(* IEC 61131-3 sources: daoli-st-library/DL_Process (part 57) *)

(* ---- FB_DL_TrapSealTrend.st ---- *)
(*
  FB_DL_TrapSealTrend  —  枕式包装封口温度随线速前馈重置 / Pillow-pack seal temperature feedforward with line-speed reset
  分类 Category : DL_Process
  码位 Code     : 16#06_0_86
  版本 Version  : 1.0.1
  溯源 Source   : Modular PID 语义借鉴 · clean-room 实现，仅借分类/参数域/命名，未复制源码
  修订 Revision : v1.0.1 (R34 终审抽检) — ① 判停改按原始线速 bSpeedStop，修正「零速保持相在曾运行后不可达」
                  （原以 fSpeedUse 判停，而 fSpeedUse 是末次有效线速替代值，恒 > 0 致 bHold 永假）；
                  ② 输入引脚 fSpeedValid 更名 bSpeedValid（BOOL 前缀红线 1，v1.0.0 无下游调用方，不构成破坏性变更）；
                  ③ 删段 7 自赋值空语句 uInfo := uInfo。接口语义与码表不变。
  功能 Function : 1) 线速前馈：封温设定 = 基准设定 + 线速偏差 × 前馈增益，线速经斜坡限速后进 PID 设定；
                  2) 线速为 0 时不得外推封温设定，改用末次有效线速并置 bHold（禁按零速反推冷设定）；
                  3) 封温设定钳到工艺窗口上下限，越限只钳位 + 报码不拒算；重置斜率须与 PID 采样周期配比，超调即判组态非法。
  边界 Boundary : ① 线速为 0 不得外推封温设定（末次有效线速 + bHold）；
                  ② 重置限速斜率与 PID 采样周期配比（每采样步进 <= fSpStepMaxC），非法即组态报码；
                  ③ 封温设定钳到工艺窗口上下限，越限只钳位 + 报码不拒算；
                  ④ 安全侧三行同向：PID 输出限 0 → 设定保持末值 → bHold 置位。
  依赖 Depends  : FB_DL_PidController（封温闭环）、FB_DL_RateLimiter（设定斜坡），均每拍无条件调用

  码表 Error codes（本件子码步进 16#10，避让邻件码位）:
    16#0002_0686 故障级：组态非法（工艺窗口上/下限倒置、增益或斜率 <= 0、采样周期 <= 0）
    16#0002_0696 故障级：前馈斜率与采样周期配比超调（单步进料过大）
    16#0002_06A6 信息级：封温设定已钳位（不置 bError，照算）
*)

TYPE E_DL_TstPhase :
(
    eIdle   := 0,   // 空闲 / Idle
    eTrack  := 10,  // 线速跟踪 / Line-speed tracking
    eHold   := 20,  // 零速保持 / Zero-speed hold
    eRun    := 30,  // 闭环调节 / Closed-loop control
    eFault  := 90   // 故障锁定 / Fault locked
);
END_TYPE

FUNCTION_BLOCK FB_DL_TrapSealTrend
VAR_INPUT
    bEnable      : BOOL;                          // 总使能，FALSE 回空闲 / Master enable
    bReset       : BOOL;                          // 复位，上升沿清故障 / Reset, clears fault
    fLineSpeedMpm: REAL;                          // 包装线速 [m/min]，域 >= 0 / Packaging line speed [m/min]
    bSpeedValid  : BOOL := TRUE;                  // 线速信号有效标志 / Line speed signal valid
    fSealTempC   : REAL;                          // 封口实测温度 [degC]，域 0~300 / Measured seal temperature [degC]
    fSealBaseC   : REAL := 150.0;                 // 基准封温设定 [degC] / Base seal temperature setpoint [degC]
    fFfGainCpm   : REAL := 0.8;                   // 线速前馈增益 [degC per m/min]，域 > 0 / Feedforward gain
    fSealWinLoC  : REAL := 120.0;                 // 工艺窗口下限 [degC] / Process window low [degC]
    fSealWinHiC  : REAL := 200.0;                 // 工艺窗口上限 [degC] / Process window high [degC]
    fSpRiseRate  : REAL := 20.0;                  // 设定上升限速 [degC/s]，域 > 0 / Setpoint rise rate [degC/s]
    fSpFallRate  : REAL := 20.0;                  // 设定下降限速 [degC/s]，域 > 0 / Setpoint fall rate [degC/s]
    fSpStepMaxC  : REAL := 5.0;                   // 单采样步进上限 [degC]，域 > 0 / Step limit per sample [degC]
    tPidSample   : TIME := T#100MS;               // PID 采样周期 [ms]，域 > 0 / PID sample period [ms]
    fKp          : REAL := 2.0;                   // 比例增益 [1] / Proportional gain
    tTi          : TIME := T#30S;                 // 积分时间 [ms] / Integral time [ms]
    tTd          : TIME := T#5S;                  // 微分时间 [ms] / Derivative time [ms]
    fEps         : REAL := 1.0E-6;                // 浮点判零容差 [1] / Floating zero tolerance
END_VAR
VAR_OUTPUT
    fSealSpC     : REAL;                          // 封温设定 [degC]，经前馈 + 限速 + 钳位 / Seal setpoint [degC]
    fPidOutPct   : REAL;                          // 加热输出 [%] / Heater output [%]
    fSpeedHold   : REAL;                          // 生效线速 [m/min]，零速时保持末次有效 / Effective line speed
    bHold        : BOOL;                          // 零速保持标志 / Zero-speed hold flag
    bClamped     : BOOL;                          // 设定钳位标志 / Setpoint clamped flag
    bError       : BOOL;                          // 故障标志，与故障级码配对 / Fault flag paired with fault codes
    uErrorId     : UDINT;                         // 事件码，0 = 无事件 / Event code, 0 = none
    eStateOut    : E_DL_TstPhase;                 // 状态机当前态，段尾单点映射 / Phase mapped at tail
END_VAR
VAR
    _eState      : E_DL_TstPhase := E_DL_TstPhase.eIdle;  // 内部状态 / Internal state
    rtrReset     : R_TRIG;                        // 复位沿 / Reset edge
    fbPid        : FB_DL_PidController;           // 封温闭环实例（无条件调用）/ Seal loop PID
    fbSpRamp     : FB_DL_RateLimiter;             // 设定斜坡实例（无条件调用）/ Setpoint ramp limiter
    bCfgOk       : BOOL;                          // 组态合法标志 / Configuration valid
    bRatioOk     : BOOL;                          // 斜率/周期配比合法 / Slope-period ratio valid
    fSpeedUse    : REAL;                          // 前馈用线速 [m/min] / Speed used for feedforward
    bSpeedStop   : BOOL;                          // 线速判停标志（按原始线速判，非替代值）/ Line stopped per raw speed
    fSpRawC      : REAL;                          // 前馈原始设定 [degC] / Raw feedforward setpoint [degC]
    fSampleS     : REAL;                          // 采样周期折算秒 [s] / Sample period in seconds
    fStepC       : REAL;                          // 单采样最大步进 [degC] / Max step per sample [degC]
    uFault       : UDINT;                         // 锁存故障码 / Latched fault code
    uInfo        : UDINT;                         // 信息级码 / Information code
END_VAR
VAR CONSTANT
    DL_TST_MSPS    : REAL := 1000.0;              // 毫秒折算秒系数 [ms/s] / Milliseconds per second
    DL_TST_TMAXC   : REAL := 300.0;               // 封温物理域上限 [degC] / Temperature domain high
END_VAR

(* === 段 0 · 实例刷新（无条件周期调用，禁入 CASE 分支）=== *)
rtrReset(CLK := bReset);                          // 每拍刷新复位沿

(* === 段 1 · 组态闸：窗口配比 / 增益正域 / 斜率-周期配比 === *)
fSampleS := TIME_TO_LREAL(tPidSample) / DL_TST_MSPS;   // 采样周期折算秒，标准转换函数
bCfgOk := (fSealWinHiC > fSealWinLoC) AND (fFfGainCpm > fEps) AND (fSpRiseRate > fEps)
          AND (fSpFallRate > fEps) AND (fSpStepMaxC > fEps) AND (fSampleS > fEps)
          AND (fSealBaseC > 0.0) AND (fSealBaseC < DL_TST_TMAXC)
          AND (fSealWinHiC = fSealWinHiC) AND (fSealWinLoC = fSealWinLoC);   // NaN 自反判据
fStepC := fSpRiseRate * fSampleS;                 // 单采样步进 = 斜率 × 周期
bRatioOk := (fStepC <= fSpStepMaxC + fEps);       // 配比闸：单步进不得超过工艺允许步进（超调即非法）
IF NOT bCfgOk THEN
    uFault := 16#0002_0686;                       // 故障级：组态非法
END_IF
IF NOT bRatioOk THEN
    uFault := 16#0002_0696;                       // 故障级：斜率与采样周期配比超调
END_IF
IF rtrReset.Q AND bCfgOk AND bRatioOk THEN
    uFault := 16#0000;                            // 复位沿清锁存（故障复位路径可达）
END_IF
uInfo := 16#0000;                                 // 信息码每拍清零

(* === 段 2 · 线速域闸：零速/无效速保持末次有效，不外推 === *)
bSpeedStop := (NOT bSpeedValid) OR (fLineSpeedMpm <> fLineSpeedMpm) OR (fLineSpeedMpm <= fEps);  // 判停只看原始线速（NaN 自反捕获）
IF NOT bSpeedStop
   AND (ABS(fLineSpeedMpm) < 1.0E6) THEN
    fSpeedUse := fLineSpeedMpm;                   // 有效线速直接采用
    fSpeedHold := fLineSpeedMpm;                  // 记入末次有效线速
ELSE
    fSpeedUse := fSpeedHold;                      // 零速/无效：用末次有效线速，禁按 0 反推
END_IF
fSpRawC := fSealBaseC + fSpeedUse * fFfGainCpm;   // 前馈原始设定 [degC]

(* === 段 3 · 设定斜坡实例（每拍无条件调用，限斜率）=== *)
fbSpRamp(bEnable := TRUE,                         // 斜坡常开
         fIn := fSpRawC,                          // 前馈原始设定
         fRateUp := fSpRiseRate,                  // 上升限速 [degC/s]
         fRateDown := fSpFallRate,                // 下降限速 [degC/s]
         bTrack := (NOT bEnable) OR (uFault <> 16#0000),   // 失能/故障：跟踪到基准设定
         fTrackValue := fSealBaseC,               // 跟踪目标 = 基准设定
         tSampleTime := tPidSample);              // 采样周期
fSealSpC := fbSpRamp.fOut;                        // 斜坡后设定

(* === 段 4 · 封温窗口钳位（越限只钳位 + 报码，不拒算）=== *)
bClamped := FALSE;                                // 钳位标志每拍重算
IF fSealSpC > fSealWinHiC THEN
    fSealSpC := fSealWinHiC;                      // 钳到上限
    bClamped := TRUE;                             // 钳位置位
    uInfo := 16#0002_06A6;                        // 信息级：设定已钳位
ELSIF fSealSpC < fSealWinLoC THEN
    fSealSpC := fSealWinLoC;                      // 钳到下限
    bClamped := TRUE;                             // 钳位置位
    uInfo := 16#0002_06A6;                        // 信息级：设定已钳位
END_IF

(* === 段 5 · 主状态机（ENUM + CASE，含 ELSE 兜底）=== *)
CASE _eState OF
E_DL_TstPhase.eIdle :
    bHold := FALSE;                               // 空闲不保持
    IF uFault <> 16#0000 THEN
        _eState := E_DL_TstPhase.eFault;          // 故障优先
    ELSIF bEnable THEN
        _eState := E_DL_TstPhase.eTrack;          // 进入跟踪相
    END_IF

E_DL_TstPhase.eTrack :
    IF bSpeedStop THEN                            // 判停按原始线速（不按前馈替代值）
        bHold := TRUE;                            // 零速：置保持，禁止外推冷设定
        _eState := E_DL_TstPhase.eHold;
    ELSE
        bHold := FALSE;                           // 有速：正常调节
        _eState := E_DL_TstPhase.eRun;
    END_IF

E_DL_TstPhase.eHold :
    bHold := TRUE;                              // 保持标志维持
    IF NOT bSpeedStop THEN
        bHold := FALSE;                          // 线速恢复即解除保持（可到达的解除路径）
        _eState := E_DL_TstPhase.eRun;
    END_IF

E_DL_TstPhase.eRun :
    IF bSpeedStop THEN                           // 判停按原始线速，与 eTrack 同源
        bHold := TRUE;                            // 线速降到 0：回保持
        _eState := E_DL_TstPhase.eHold;
    ELSIF NOT bEnable THEN
        _eState := E_DL_TstPhase.eIdle;           // 失能回空闲
    ELSIF uFault <> 16#0000 THEN
        _eState := E_DL_TstPhase.eFault;          // 故障拦截
    END_IF

E_DL_TstPhase.eFault :
    bHold := TRUE;                                // 故障态保持（安全侧）
    IF uFault = 16#0000 THEN
        _eState := E_DL_TstPhase.eIdle;           // 解锁回空闲
    END_IF

ELSE
    _eState := E_DL_TstPhase.eFault;              // 非法状态拦截
    uFault := 16#0002_0686;                       // 故障级：相 ID 越界（枚举兜底路径）
END_CASE

(* === 段 6 · 封温闭环实例（每拍无条件调用）=== *)
fbPid(bEnable := bEnable AND (NOT bHold) AND (uFault = 16#0000),   // 保持/故障时禁调节
      bManual := FALSE,                           // 自动模式
      fManualValue := 0.0,                        // 手动值未用
      fSetpoint := fSealSpC,                      // 设定 = 钳位后封温
      fActual := fSealTempC,                      // 实测封温
      fKp := fKp,                                 // 比例增益
      tTi := tTi,                                 // 积分时间
      tTd := tTd,                                 // 微分时间
      fDeadband := 0.5,                           // 控制死区 [degC]，防抖
      bIncremental := FALSE,                      // 位置式
      rOutMin := 0.0,                             // 输出下限 0%（安全侧）
      rOutMax := 100.0,                           // 输出上限 100%
      tSampleTime := tPidSample,                  // 采样周期
      bTrack := bHold OR (uFault <> 16#0000),     // 保持/故障：跟踪 0 输出
      fTrackValue := 0.0,                         // 跟踪值 0（断加热）
      bReset := rtrReset.Q);                      // 复位沿清积分

(* === 段 7 · 输出映射（安全三行同向）=== *)
IF bHold OR (uFault <> 16#0000) THEN
    fPidOutPct := 0.0;                            // 保持/故障：加热输出 0（驱动方向安全）
    bHold := TRUE;                                // 保持判据与输出同向（设定同步冻结在段 3/4 末值）
ELSE
    fPidOutPct := fbPid.fOut;                     // 正常：取 PID 输出
END_IF
IF NOT bEnable THEN
    fPidOutPct := 0.0;                            // 失能输出 0
END_IF
bError := (uFault <> 16#0000);                    // 故障标志仅由故障级码置位（R45 配对）
IF bError THEN
    uErrorId := uFault;                           // 故障级优先上报
ELSE
    uErrorId := uInfo;                            // 否则上报信息级码
END_IF
eStateOut := _eState;                             // 输出枚举段尾单点映射（N2 规则）
END_FUNCTION_BLOCK

(* ---- FB_DL_TrayerNestingCtrl.st ---- *)
(*==============================================================================
 * 组件名称 (Component)  : FB_DL_TrayerNestingCtrl
 * 所属子库 (Sublibrary) : DL_Process
 * 当前版本 (Version)    : 1.0.0
 * 兼容性   (Platform)   : CODESYS 3.5+ / TwinCAT 3 / 汇川 InoProShop / 施耐德 Machine Expert
 *                         仅依赖 Standard.library（R_TRIG），零厂商私有库
 * 功能描述 (Function)   : 电芯托盘堆叠嵌套调度（层 × 列网格占位）。
 *                         按"层从下往上、列从左往右"的蛇形无关直线序逐格占位；每来一颗电芯占一格，
 *                         列到边界回卷到下一层首列；**NG 通道避让**：某一列指定为 NG 列时，
 *                         该列在每一层都被整体跳过（整列不占位、不计入容量）；
 *                         合法格占满即判"栈满"并锁存 bTrayFull，等待取盘沿（bTrayTaken）或复位沿解除。
 *                         **语义复用（非实例复用）**：本件按 R47 批次"批内零 .st 文件级依赖"纪律，
 *                         不实例化 FB_DL_LifoStack，而是复用其三条已固化语义——
 *                         ① 入栈前判满、满则拒入并锁存；② 出栈仅由显式"取走"沿触发；
 *                         ③ 满/空判定以计数与容量比较为准，不以指针相等为准。
 *                         验收向量：
 *                           ① 3 层 × 4 列、NG 列 = 2 → 容量 = 3×(4−1) = 9 格
 *                           ② 2 层 × 2 列、NG 列 = 1 → 容量 = 2×(2−1) = 2 格
 *                           ③ 2 层 × 2 列、NG 列 = 0 → 容量 = 4 格
 *                           ④ 任一层列数 = 0 → 组态非法锁存，不进入占位
 * 接口     (Interface)  : 入 bStart 启动沿、bTrayTaken 取盘沿（解除栈满）、iLayerCnt 层数、iColCnt 列数、
 *                         iNgCol 避让列号（1 基，0 = 无）、bCellPresent 电芯到位沿、bPlaceAllowed 上料允许
 *                         （外部互锁）、bReset 故障复位沿；
 *                         出 iLayerOut / iColOut 当前待占格坐标（1 基）、bPlaceCmd 占位脉冲（单拍）、
 *                         bLayerDone 换层脉冲（单拍）、bTrayFull 栈满锁存、iPlacedCnt 已占格数、
 *                         bNgSkipped 当拍发生 NG 列跳过、eState 相、eCause 成因、bError 故障标志。
 * 边界     (Boundary)   : ① **属主边界（写死）：本件只算"下一颗电芯放哪一格"，不驱动吸盘/夹具/
 *                         升降台伺服**；取放动作由执行件（I_DL_Cylinder 族 / 运动件）承担；
 *                         ② **网格组态闸**：层数或列数 ≤ 0 或超上限（100×100）→ 锁存 eCfgIllegal，
 *                         不进入占位（零容量网格会让"栈满"永假，属静默失效 R179）；
 *                         ③ **NG 列域闸**：iNgCol 越界（<0 或 > 列数）→ 锁存 eCfgIllegal；
 *                         ④ **索引越界钳位**：前进循环带 _uGuard 计数器（上界 = 总格数 + 列数 + 2），
 *                         循环必然收敛，绝不靠"数据一定合法"保证终止；
 *                         ⑤ eFault 可迁出：bReset 上升沿 → eIdle（解除式自证：bReset 为外部引脚，
 *                         不受任何锁存量门控，恒可达）；
 *                         ⑥ 零全局耦合、零物理地址。
 * 分工声明 (Scope)      : 本件只管"托盘格位调度与栈满判定"。不接管：电芯取放动作时序（顺控件）、
 *                         NG 电芯的下游分选（分选件）、托盘身份绑定（RFID 件）。
 * 来源标签 (Source Tag) : ROADMAP 空勾真缺口 P2（托盘嵌套调度，自研 clean-room）
 * 码表     (Codes)      : 本件不占用任何全局数字码位（零码位范式 R297）；诊断由 BOOL + ENUM 出口承担。
 * 红线自检 (Redline)    : R1 ✓ 零 GVL/VAR_EXTERNAL ｜ R2 ✓ 零 %I/%Q/%M ｜ R3 ✓ 纯 IEC 61131-3
 *                         R4 ✓ 组态双闸 + 循环计数器 + 索引钳位 ｜ R5 ✓ 声明逐行同行双语注释
 *                         R6 ✓ ENUM+CASE 含 ELSE 兜底 ｜ R7 ✓ R_TRIG 段 0 无条件刷新（本件无 TON）
 * 修订历史 (Revision)   : 2026-11-19  v1.0.0  R47 首版（批次 1 · 序号 4）
 *==============================================================================*)

TYPE E_DL_TncState :
(
    eIdle  := 0,    // 待机相（等启动或等取盘） / Idle, awaiting start or tray removal
    eNest  := 10,   // 占位相（逐颗占格） / Nesting, one cell per cell-in
    eFull  := 20,   // 栈满相（锁存等取盘） / Full, latched awaiting tray removal
    eFault := 90    // 故障相（等复位） / Fault, awaiting reset
);
END_TYPE

TYPE E_DL_TncCause :
(
    eNone      := 0,   // 无异常 / No anomaly
    eCfgIllegal:= 1,   // 组态非法（层数/列数/NG 列越域） / Illegal grid configuration
    eFullNoCell    := 2,   // 栈满后仍有电芯到位（拒入） / Cell arrived while full, rejected
    eRejectNoPermit:= 3,   // 上料允许缺失致电芯被拒 / Cell rejected, place permit absent
    ePhaseBad      := 4    // 非法相位兜底 / Illegal phase fallback
);
END_TYPE

FUNCTION_BLOCK FB_DL_TrayerNestingCtrl
VAR_INPUT
    bStart       : BOOL := FALSE;   // 启动沿，进入占位相 [-] / Start edge, enters nesting
    bTrayTaken   : BOOL := FALSE;   // 取盘沿，解除栈满并清零计数 [-] / Tray-removed edge, clears the full latch
    iLayerCnt    : INT := 1;        // 层数，域 1..100 [层] / Layer count, domain 1..100
    iColCnt      : INT := 1;        // 每层列数，域 1..100 [列] / Columns per layer, domain 1..100
    iNgCol       : INT := 0;        // NG 避让列号（1 基；0 = 不避让） [列] / NG column index, 1-based, 0 = none
    bCellPresent : BOOL := FALSE;   // 电芯到位信号（上升沿占一格） [-] / Cell-present signal, rising edge takes one cell
    bPlaceAllowed: BOOL := FALSE;   // 上料允许（外部互锁，FALSE 时拒占位） [-] / Place permit from the external interlock
    bReset       : BOOL := FALSE;   // 故障复位沿 [-] / Fault reset edge
END_VAR
VAR_OUTPUT
    iLayerOut  : INT := 0;                  // 当前待占格所在层（1 基） [层] / Current target layer, 1-based
    iColOut    : INT := 0;                  // 当前待占格所在列（1 基） [列] / Current target column, 1-based
    bPlaceCmd  : BOOL := FALSE;             // 占位脉冲，单拍 [-] / Place command, single-scan pulse
    bLayerDone : BOOL := FALSE;             // 换层脉冲，单拍 [-] / Layer-change pulse, single-scan
    bTrayFull  : BOOL := FALSE;             // 栈满锁存（等取盘或复位） [-] / Tray full, latched
    iPlacedCnt : INT := 0;                  // 已占格数 [格] / Occupied cell count
    bNgSkipped : BOOL := FALSE;             // 当拍发生过 NG 列跳过 [-] / An NG column was skipped this scan
    eState     : E_DL_TncState := E_DL_TncState.eIdle;   // 相出口 [-] / Phase outlet
    eCause     : E_DL_TncCause := E_DL_TncCause.eNone;   // 成因出口（R190 归因唯一） [-] / Cause outlet
    bError     : BOOL := FALSE;             // 故障标志 [-] / Error flag
END_VAR
VAR
    _eState    : E_DL_TncState := E_DL_TncState.eIdle;   // 内部相（CASE 唯一写入目标） / Internal phase
    _eCause    : E_DL_TncCause := E_DL_TncCause.eNone;   // 成因锁存量 / Latched cause
    _bFault    : BOOL := FALSE;             // 故障锁存位 / Latched fault bit
    _bFull     : BOOL := FALSE;             // 栈满锁存位（与 bTrayFull 同源） / Latched full bit
    _iLayer    : INT := 1;                  // 内部层指针（1 基） / Internal layer cursor
    _iCol      : INT := 1;                  // 内部列指针（1 基） / Internal column cursor
    _iPlaced   : INT := 0;                  // 内部已占格计数 / Internal occupied counter
    _iCap      : INT := 0;                  // 本盘合法格容量（不含 NG 列） / Legal capacity excluding the NG column
    _bPlaceCmd : BOOL := FALSE;             // 占位脉冲内部位（单拍） / Internal place pulse
    _bLayerDone: BOOL := FALSE;             // 换层脉冲内部位（单拍） / Internal layer-change pulse
    _bNgSkipped: BOOL := FALSE;             // NG 跳过内部位（单拍） / Internal NG-skip flag
    _bCfgBad   : BOOL := FALSE;             // 组态非法当拍量 / Illegal configuration this scan
    _bAdvDone  : BOOL := FALSE;             // 前进循环收敛标志 / Advance-loop convergence flag
    _uGuard    : UINT := 0;                 // 前进循环计数器（防死循环） / Advance-loop guard counter
    rtStart    : R_TRIG;                    // 启动沿实例，段 0 无条件调用 / Start edge instance
    rtReset    : R_TRIG;                    // 复位沿实例，段 0 无条件调用 / Reset edge instance
    rtTaken    : R_TRIG;                    // 取盘沿实例，段 0 无条件调用 / Tray-removed edge instance
    rtCell     : R_TRIG;                    // 电芯到位沿实例，段 0 无条件调用 / Cell-present edge instance
END_VAR
VAR CONSTANT
    DL_TNC_MAX_LAYER : INT := 100;          // 层数上限（超限判组态非法） [层] / Layer upper bound
    DL_TNC_MAX_COL   : INT := 100;          // 列数上限（超限判组态非法） [列] / Column upper bound
    DL_TNC_GUARD_MAX : UINT := 20002;       // 前进循环守护上限（100×100 + 100 + 2） [次] / Advance guard limit
END_VAR

(* —— 段 0：组态闸 + 四枚沿实例无条件周期刷新（R228A） —— *)
_bCfgBad := (iLayerCnt <= 0) OR (iLayerCnt > DL_TNC_MAX_LAYER)          // 层数须在 1..100 / Layer count within 1..100
         OR (iColCnt <= 0) OR (iColCnt > DL_TNC_MAX_COL)                // 列数须在 1..100 / Column count within 1..100
         OR (iNgCol < 0) OR (iNgCol > iColCnt);                          // NG 列号须为 0 或落在列域内 / NG index within the column domain
rtStart(CLK := bStart);                                                  // 启动沿 / Start edge
rtReset(CLK := bReset);                                                  // 复位沿 / Reset edge
rtTaken(CLK := bTrayTaken);                                              // 取盘沿 / Tray-removed edge
rtCell(CLK := bCellPresent);                                             // 电芯到位沿 / Cell-present edge

(* —— 段 1：单拍量预清零（锁存量 _eCause/_bFault/_iPlaced 不入清单，R107） —— *)
_bPlaceCmd  := FALSE;                                                    // 占位脉冲预清 / Place pulse preset
_bLayerDone := FALSE;                                                    // 换层脉冲预清 / Layer pulse preset
_bNgSkipped := FALSE;                                                    // NG 跳过标志预清 / NG-skip preset
bError      := FALSE;                                                    // 故障标志预清（R45 配对） / Error preset

(* —— 段 2：组态闸（非法即锁存，不进入占位） —— *)
IF _bCfgBad THEN
    _bFault := TRUE;                                                     // 锁存 / Latch
    _eCause := E_DL_TncCause.eCfgIllegal;                                // 归因：组态非法 / Cause: illegal configuration
    _eState := E_DL_TncState.eFault;                                     // 入故障相 / Enter fault phase
END_IF

(* —— 段 3：迁出链与取盘链（两条出口显式写出，R228B） —— *)
IF rtReset.Q THEN
    _bFault  := FALSE;                                                   // 清故障锁存 / Clear fault latch
    _bFull   := FALSE;                                                   // 清栈满锁存 / Clear full latch
    _eCause  := E_DL_TncCause.eNone;                                     // 清成因 / Clear cause
    _iPlaced := 0;                                                       // 计数清零 / Clear the counter
    _iLayer  := 1;                                                       // 层指针回 1 / Layer cursor back to 1
    _iCol    := 1;                                                       // 列指针回 1 / Column cursor back to 1
    _eState  := E_DL_TncState.eIdle;                                     // 回待机相 / Back to idle
END_IF
IF rtTaken.Q AND (_eState <> E_DL_TncState.eFault) THEN
    _bFull   := FALSE;                                                   // 取盘解除栈满 / Tray removal clears the full latch
    _iPlaced := 0;                                                       // 计数清零 / Clear the counter
    _iLayer  := 1;                                                       // 层指针回 1 / Layer cursor back to 1
    _iCol    := 1;                                                       // 列指针回 1 / Column cursor back to 1
    _eState  := E_DL_TncState.eIdle;                                     // 回待机相 / Back to idle
END_IF

(* —— 段 4：容量计算（总格数 − NG 列整列格数；组态合法时恒 ≥ 0） —— *)
IF NOT _bCfgBad THEN
    _iCap := iLayerCnt * iColCnt;                                        // 总格数 / Total cells
    IF iNgCol > 0 THEN
        _iCap := _iCap - iLayerCnt;                                      // 扣除 NG 列整列 / Deduct the whole NG column
    END_IF
END_IF

(* —— 段 5：相迁移（只在无故障时推进；每相出口条件显式成对） —— *)
IF (NOT _bFault) AND (NOT _bCfgBad) THEN
    CASE _eState OF

    E_DL_TncState.eIdle:
        IF rtStart.Q THEN
            _iLayer := 1;                                                // 层指针首层 / First layer
            IF (iNgCol = 1) AND (iColCnt >= 2) THEN
                _iCol := 2;                                              // 首列即 NG：起始列右移一格 / First column is NG, start at column 2
            ELSE
                _iCol := 1;                                              // 否则首列起步 / Otherwise start at column 1
            END_IF
            _iPlaced := 0;                                               // 计数清零 / Counter cleared
            _eState := E_DL_TncState.eNest;                              // 进占位相 / Enter nesting
        END_IF

    E_DL_TncState.eNest:
        IF rtCell.Q AND bPlaceAllowed THEN
            _bPlaceCmd := TRUE;                                          // 占位脉冲（内部位，段 7 单点映射） / Internal place pulse
            _iPlaced := _iPlaced + 1;                                    // 占位计数 +1 / Increment the counter

            (* 前进到下一合法格：列 +1，越界回卷到下一层首列，NG 列整体跳过 *)
            _uGuard  := 0;                                               // 守护计数器归零 / Guard reset
            _bAdvDone:= FALSE;                                           // 收敛标志复位 / Convergence flag reset
            WHILE (NOT _bAdvDone) AND (_uGuard < DL_TNC_GUARD_MAX) DO
                _uGuard := _uGuard + 1;                                  // 计数器推进 / Guard advance
                _iCol := _iCol + 1;                                      // 列前进一格 / Column step
                IF _iCol > iColCnt THEN
                    _iCol := 1;                                          // 列回卷 / Column wrap
                    _iLayer := _iLayer + 1;                              // 换层 / Next layer
                    _bLayerDone := TRUE;                                 // 换层脉冲（内部位） / Internal layer pulse
                END_IF
                IF _iLayer > iLayerCnt THEN
                    _bAdvDone := TRUE;                                   // 层耗尽：指针停（不再寻格） / Layers exhausted
                ELSIF (iNgCol > 0) AND (_iCol = iNgCol) THEN
                    _bNgSkipped := TRUE;                                 // NG 列：跳过并继续寻格 / NG column skipped, keep seeking
                ELSE
                    _bAdvDone := TRUE;                                   // 找到合法格 / Legal cell found
                END_IF
            END_WHILE

            IF _iPlaced >= _iCap THEN
                _bFull   := TRUE;                                        // 栈满锁存（入栈前判满语义） / Full latch, pre-push check
                _eState  := E_DL_TncState.eFull;                         // 进栈满相 / Enter full phase
            END_IF
        ELSIF rtCell.Q AND (NOT bPlaceAllowed) THEN
            _eCause := E_DL_TncCause.eRejectNoPermit;                    // 归因：互锁未放开致电芯被拒 / Cause: cell rejected, permit absent
        END_IF

    E_DL_TncState.eFull:
        IF rtCell.Q THEN
            _eCause := E_DL_TncCause.eFullNoCell;                        // 满盘期电芯到位：拒入并留痕 / Cell during full: rejected and recorded
        END_IF

    E_DL_TncState.eFault:
        ;                                                                // 故障相：由段 3 复位沿迁出 / Exit handled by the reset edge in stage 3

    ELSE
        _eCause := E_DL_TncCause.ePhaseBad;                              // 归因：非法相位 / Cause: illegal phase
        _bFault := TRUE;                                                 // 锁存 / Latch
        _eState := E_DL_TncState.eFault;                                 // 强拉故障相 / Force fault phase

    END_CASE
END_IF

(* —— 段 6：栈满与故障的交汇（满盘后故障优先展示，满锁存保持） —— *)
IF _bFull AND (_eState = E_DL_TncState.eNest) THEN
    _eState := E_DL_TncState.eFull;                                      // 满锁存与相对齐 / Align the phase with the full latch
END_IF

(* —— 段 7：出口单点映射（名实双出口，R191） —— *)
iLayerOut  := _iLayer;                                                   // 待占层层号 / Target layer
iColOut    := _iCol;                                                     // 待占格列号 / Target column
bPlaceCmd  := _bPlaceCmd;                                                // 占位脉冲单拍出口 / Place pulse outlet
bLayerDone := _bLayerDone;                                               // 换层脉冲单拍出口 / Layer pulse outlet
bNgSkipped := _bNgSkipped;                                               // NG 跳过标志出口 / NG-skip outlet
bTrayFull  := _bFull;                                                    // 栈满出口 / Full outlet
iPlacedCnt := _iPlaced;                                                  // 已占格数出口 / Occupied count outlet
eState     := _eState;                                                   // 相出口 / Phase outlet
eCause     := _eCause;                                                   // 成因出口 / Cause outlet
bError     := _bFault OR _bCfgBad;                                       // 故障标志 = 锁存或组态非法 / Error = latch or illegal config

END_FUNCTION_BLOCK

(* ---- FB_DL_TrayLoadVacuum.st ---- *)
(*==============================================================================
 * 组件名称 (Component)  : FB_DL_TrayLoadVacuum
 * 所属子库 (Sublibrary) : DL_Process
 * 当前版本 (Version)    : 1.0.0
 * 兼容性 (Platform)     : CODESYS 3.5+ / TwinCAT 3 / 汇川 InoProShop / 施耐德 Machine Expert
 *                         仅依赖 Standard.library（TON / TOF / R_TRIG / F_TRIG），零厂商私有库
 * 功能描述 (Function)   : 电池片花篮真空取放顺控。吸取相开真空阀，真空反馈
 *                         在 tVacOnDelay 内不到达即吸取超时故障（独立成因）；
 *                         放片相关真空并以 TOF 定宽输出破真空吹气脉冲
 *                         （宽度 tBlowWidth + 1 扫描拍，头注释明示），吹气
 *                         结束沿收口 bPlaceDone。与 VacuumEjector（真空发生
 *                         设备件）分工：本件是取放顺控中破真空定宽脉冲的
 *                         时序件。
 * 来源标签 (Origin)     : ROADMAP §9.3 P2（L418），自研 clean-room
 * 边界语义 (Boundary)   : ① 吸取超时 TON 电平计时（非自复位周期窗）；
 *                         ② 吹气定宽用 TOF（触发单拍 → 展宽 tBlowWidth），
 *                         结束沿用 F_TRIG（段 0 无条件刷新）；
 *                         ③ 故障相真空阀强制关断（安全侧失真空）；
 *                         ④ 组态闸：两时间量正域 → 故障锁存。
 * 输出语义 (Fallback)   : 【R191】bEnable = FALSE → 双阀输出强制 FALSE（阀类
 *                         出口失能必须收敛）；eFault 相 → 真空阀 FALSE +
 *                         bError = TRUE。
 * 码位     (Codes)      : 按 R297 范式零 16# 码位硬编码；错误出口 BOOL+ENUM(eCause)。
 * 红线自检 (Redline)    : 7 项红线已自检：R1 零全局 ✓｜R2 零物理地址 ✓｜R3 纯 IEC ✓
 *                         R4 除零无涉/组态闸 ✓｜R5 双语同行注释 ✓
 *                         R6 CASE 带 ELSE 兜底迁 eFault ✓｜R7 TON/TOF/R_TRIG/F_TRIG 段 0 无条件刷新 ✓
 * 验收向量 (Acceptance) : V1 取片申请沿 → 真空阀 TRUE，bVacFb 在 tVacOnDelay
 *                         内到达 → bPickDone 单拍进保持相；
 *                         V2 反馈超 tVacOnDelay 未到 → eVacFail 故障锁存，
 *                         真空阀关断；
 *                         V3 放片申请沿 → 真空阀关 + 吹气阀展宽 tBlowWidth
 *                         后 bPlaceDone 单拍回待机。
 * 修订历史 (Revision)   : 2026-11-20  v1.0.0  R51 首版（批 4 · 序号 16）
 *==============================================================================*)
TYPE E_DL_TlvState :
(
    eIdle  := 0,                             (* 待机（双阀关） / Idle *)
    ePick  := 10,                            (* 真空吸取 / Vacuum pick *)
    eHold  := 20,                            (* 吸取保持（待放片申请） / Hold *)
    ePlace := 30,                            (* 破真空吹气放片 / Blow-off place *)
    eFault := 90                             (* 故障锁存相 / Fault latched phase *)
);
END_TYPE

TYPE E_DL_TlvCause :
(
    eNone     := 0,                          (* 无故障成因 / No cause *)
    eCfgIllegal := 1,                        (* 组态非法：时间量越域 / Illegal config *)
    eVacFail  := 2,                          (* 吸取真空反馈超时 / Vacuum feedback timeout *)
    ePhaseBad := 3                           (* 非法相位兜底 / Illegal phase fallback *)
);
END_TYPE

FUNCTION_BLOCK FB_DL_TrayLoadVacuum
VAR_INPUT
    bPickReq   : BOOL := FALSE;              (* 取片申请沿 [-] / Pick request edge *)
    bPlaceReq  : BOOL := FALSE;              (* 放片申请沿 [-] / Place request edge *)
    bVacFb     : BOOL := FALSE;              (* 真空到达反馈电平 [-] / Vacuum feedback level *)
    tVacOnDelay: TIME := T#2S;               (* 真空建立超时，域 > T#0S [ms] / Vacuum build timeout *)
    tBlowWidth : TIME := T#500MS;            (* 破真空吹气定宽，域 > T#0S [ms] / Blow pulse width *)
    bEnable    : BOOL := TRUE;               (* 使能 [-] / Enable *)
    bReset     : BOOL := FALSE;              (* 复位命令，上升沿清全部 [-] / Reset command *)
END_VAR
VAR_OUTPUT
    bVacValve  : BOOL;                       (* 真空阀输出 [-] / Vacuum valve outlet *)
    bBlowValve : BOOL;                       (* 破真空吹气阀输出（定宽脉冲）[-] / Blow valve outlet *)
    bPickDone  : BOOL;                       (* 吸取完成单拍位 [-] / Pick-done pulse *)
    bPlaceDone : BOOL;                       (* 放片完成单拍位 [-] / Place-done pulse *)
    nCycleCnt  : UDINT;                      (* 累计取放循环数 [次] / Cycle count *)
    eState     : E_DL_TlvState;              (* 状态出口 / State outlet *)
    eCause     : E_DL_TlvCause;              (* 故障成因出口 / Fault cause outlet *)
    bError     : BOOL;                       (* 故障锁存标志 [-] / Fault latch flag *)
END_VAR
VAR
    _eState   : E_DL_TlvState := E_DL_TlvState.eIdle;     (* 内部相位（CASE 唯一写入目标） / Internal phase *)
    _eCause   : E_DL_TlvCause := E_DL_TlvCause.eNone;     (* 故障成因锁存量 / Latched cause *)
    rtPick    : R_TRIG;                      (* 取片沿实例，段 0 无条件调用 / Pick edge instance *)
    rtPlace   : R_TRIG;                      (* 放片沿实例，段 0 无条件调用 / Place edge instance *)
    rtReset   : R_TRIG;                      (* 复位沿实例，段 0 无条件调用 / Reset edge instance *)
    tonVac    : TON;                         (* 真空建立超时计时，段 0 无条件调用 / Vacuum timeout timer *)
    toBlow    : TOF;                         (* 吹气定宽展宽（TOF 下降沿后保持 PT）[ms] / Blow width stretcher *)
    ftBlow    : F_TRIG;                      (* 吹气结束沿实例，段 0 无条件调用 / Blow-end edge instance *)
    _bVacOn   : BOOL;                        (* 真空阀指令锁存 [-] / Vacuum valve latch *)
    _bBlowFire: BOOL;                        (* 吹气触发单拍量（TOF 输入）[-] / Blow fire pulse *)
    _bBlowAct : BOOL;                        (* 吹气进行中锁存（结束沿判据）[-] / Blow-active latch *)
    _nCycles  : UDINT;                       (* 循环计数锁存 [次] / Cycle count latch *)
    _bPickD   : BOOL;                        (* 吸取完成单拍量 [-] / Pick-done work *)
    _bPlaceD  : BOOL;                        (* 放片完成单拍量 [-] / Place-done work *)
    _bFault   : BOOL;                        (* 故障锁存位 / Latched fault bit *)
    _bCfgBad  : BOOL;                        (* 组态非法当拍量 / Illegal config this scan *)
END_VAR

(* —— 段 0：当拍判据派生 + 实例无条件刷新（R228A） —— *)
_bCfgBad := (tVacOnDelay <= T#0S) OR (tBlowWidth <= T#0S);   (* 组态闸（R151 全引脚） / Config gate *)
rtPick(CLK := bPickReq);                     (* 取片沿每拍必调 / Pick edge every scan *)
rtPlace(CLK := bPlaceReq);                   (* 放片沿每拍必调 / Place edge every scan *)
rtReset(CLK := bReset);                      (* 复位沿每拍必调 / Reset edge every scan *)
tonVac(IN := (_eState = E_DL_TlvState.ePick) AND (NOT bVacFb), PT := tVacOnDelay);   (* 真空建立超时（电平计时非周期窗） / Vacuum timeout *)
toBlow(IN := _bBlowFire, PT := tBlowWidth);  (* 吹气展宽：单拍触发 → Q 保持 tBlowWidth（输出脉宽 = PT + 1 拍，头注释明示） / Blow stretcher *)
ftBlow(CLK := toBlow.Q);                     (* 吹气结束沿每拍必调 / Blow-end edge every scan *)

(* —— 段 1：单拍量预清零（R107） —— *)
_bBlowFire := FALSE;                         (* 吹气触发预清，唯一分支置位 / Blow fire preset *)
_bPickD := FALSE;                            (* 吸取完成预清 / Pick-done preset *)
_bPlaceD := FALSE;                           (* 放片完成预清 / Place-done preset *)
bPickDone := FALSE;                          (* 吸取完成出口预清 / Pick-done outlet preset *)
bPlaceDone := FALSE;                         (* 放片完成出口预清 / Place-done outlet preset *)

(* —— 段 2：复位沿处理（作用域：清故障 + 清阀锁存 + 清吹气锁存 + 清计数 + 迁 eIdle，R283 逐项声明） —— *)
IF rtReset.Q THEN
    _bFault := FALSE;                        (* 清故障锁存 / Clear fault *)
    _eCause := E_DL_TlvCause.eNone;          (* 清成因 / Clear cause *)
    _bVacOn := FALSE;                        (* 清真空阀锁存 / Clear valve latch *)
    _bBlowAct := FALSE;                      (* 清吹气锁存 / Clear blow latch *)
    _nCycles := 0;                           (* 清循环计数 / Clear count *)
    _eState := E_DL_TlvState.eIdle;          (* 迁待机相 / Back to idle *)
END_IF

(* —— 段 3：组态闸故障锁存（R45 配对；锁存至复位沿，R189） —— *)
IF _bCfgBad AND NOT _bFault THEN
    _bFault := TRUE;                         (* 锁存故障位 / Latch fault *)
    _eCause := E_DL_TlvCause.eCfgIllegal;    (* 成因：组态非法 / Cause: illegal config *)
    _eState := E_DL_TlvState.eFault;         (* 同步迁故障相 / Migrate to fault *)
END_IF

(* —— 段 4：CASE 主状态机（ELSE 兜底迁 eFault，红线 6） —— *)
CASE _eState OF
    E_DL_TlvState.eIdle:                     (* 待机相 / Idle *)
        IF rtPick.Q AND bEnable AND (NOT _bFault) THEN
            _bVacOn := TRUE;                 (* 开真空阀 / Open vacuum valve *)
            _eState := E_DL_TlvState.ePick;  (* 进入吸取 / Enter pick *)
        END_IF
    E_DL_TlvState.ePick:                     (* 吸取相：等真空反馈或超时 / Pick *)
        IF bVacFb THEN                       (* 反馈到达：吸取完成（过渡态三段：本拍发完成脉冲并迁相/下拍预清，R80） / Feedback arrived *)
            _bPickD := TRUE;                 (* 内部完成量置位（统一出口映射单拍，R189 两段式） / Internal done set *)
            _eState := E_DL_TlvState.eHold;  (* 进保持相 / Enter hold *)
        ELSIF tonVac.Q THEN                  (* 建立超时：故障锁存（R190 独立成因） / Build timeout *)
            _eCause := E_DL_TlvCause.eVacFail;   (* 成因：真空超时 / Cause: vac timeout *)
            _bFault := TRUE;                 (* 故障锁存（R45 配对） / Latch fault *)
            _bVacOn := FALSE;                (* 故障相真空阀关断（安全侧，边界③） / Close valve safe side *)
            _eState := E_DL_TlvState.eFault; (* 迁故障相 / To fault *)
        END_IF
    E_DL_TlvState.eHold:                     (* 保持相：待放片申请 / Hold *)
        IF rtPlace.Q AND bEnable AND (NOT _bFault) THEN
            _bVacOn := FALSE;                (* 关真空阀（破真空） / Close vacuum valve *)
            _bBlowFire := TRUE;              (* 吹气触发单拍（TOF 展宽定宽） / Fire blow pulse *)
            _bBlowAct := TRUE;               (* 置吹气进行锁存 / Set blow-active *)
            _eState := E_DL_TlvState.ePlace; (* 进放片相 / Enter place *)
        END_IF
    E_DL_TlvState.ePlace:                    (* 放片相：吹气定宽至结束沿 / Place *)
        IF ftBlow.Q AND _bBlowAct THEN       (* 吹气结束沿：收口（过渡态三段：本拍发单拍/下拍预清，R80） / Blow-end edge: close out *)
            _bBlowAct := FALSE;              (* 清吹气锁存 / Clear blow latch *)
            _bPlaceD := TRUE;                (* 内部完成量置位 / Internal done set *)
            _nCycles := _nCycles + 1;        (* 循环计数（UDINT 回绕工程安全） / Count cycle *)
            _eState := E_DL_TlvState.eIdle;  (* 回待机 / Back to idle *)
        END_IF
    E_DL_TlvState.eFault:                    (* 故障相：阀已安全关断，仅复位沿出 / Fault *)
        ;                                    (* 锁存回放（R28） / Replay from latch *)
    ELSE                                     (* 非法相位兜底迁安全态 / Illegal phase fallback *)
        _eState := E_DL_TlvState.eFault;     (* 迁故障相 / To fault *)
        _bFault := TRUE;                     (* 同步锁存 / Latch *)
        _eCause := E_DL_TlvCause.ePhaseBad;  (* 成因：非法相位 / Cause: illegal phase *)
END_CASE

(* —— 段 5：出口映射（完成脉冲两段式统一出口，R189；阀出口与状态同源 R191） —— *)
bPickDone := _bPickD;                        (* 吸取完成单拍出口 / Pick-done outlet *)
bPlaceDone := _bPlaceD;                      (* 放片完成单拍出口 / Place-done outlet *)
bVacValve := _bVacOn AND bEnable AND (NOT _bFault);   (* 真空阀出口（失能/故障收敛 FALSE） / Vacuum valve outlet *)
bBlowValve := toBlow.Q AND _bBlowAct AND bEnable AND (NOT _bFault);   (* 吹气阀出口（定宽 + 门控收敛） / Blow valve outlet *)
nCycleCnt := _nCycles;                       (* 循环计数出口 / Count outlet *)
bError := _bFault;                           (* 故障标志镜像 / Fault flag mirror *)
eState := _eState;                           (* 状态出口 / State outlet *)
eCause := _eCause;                           (* 成因出口 / Cause outlet *)
END_FUNCTION_BLOCK

(* ---- FB_DL_TrayMonthRotate.st ---- *)
(*
  ==================================================================
  组件名 Component  : FB_DL_TrayMonthRotate
  分类   Category   : DL_Process
  版本   Version    : 1.0.0
  功能   Purpose    : 托盘月度轮换保养排程。按「上次保养月」与保养周期（月数）逐盘
                      判到期，到期盘打包成 12 位到期掩码字，并给本月轮换优先盘号
                      （按月份在托盘序列上轮转），支持保养完成脉冲回写上次保养月。
  溯源   Origin     : 月度轮换保养为通用设备维护排程语义；本件为 clean-room 实现，
                      仅借鉴来源分类与参数域组织（来源标签 roadmap-p2-tray），
                      道莅原创设计，未复制任何闭源代码行。
  平台   Platform   : 纯 IEC 61131-3（WORD / SHL / MOD / R_TRIG，无私有库）
  作者   Author     : 道莅代码库 · PLC 编程专家（R55）
  ------------------------------------------------------------------
  边界 Boundary     :
                      一 本件只出到期掩码与优先盘号，不启动保养动作、不判保养质量；
                      二 周期判据按月数差计，跨年回绕按「月差加 12」补齐，只覆盖一周年内；
                      三 保养完成回写由 bMaintDone 上升沿 + nMaintTray 触发，
                         托盘号经回钳 1..12 后写入调用方持有的上次保养月表；
                      四 未保养盘（上次保养月小于 1）一律立即到期，不参与月差计算；
                      五 无全局变量、无外部变量声明、无物理地址寻址。
  输出契约 Output contract:
                      wDueMask 位 i-1 对应托盘 i，自证向量：仅 1 号盘到期 → 16#0001，
                      仅 12 号盘到期 → 16#0800；
                      nPriTray 为 1..nTrayCount 内的轮换优先盘号，该盘到期时 bPriDue 为真；
                      eCause 故障级成因与 bError 配对（R45），信息级永不置 bError。
  修订记录 Revision  :
    2026-11-20  v1.0.0  R55 首版（批 2 · 序号 7）
  ==================================================================
*)

TYPE E_DL_TmrCause :
(
    eNone       := 0,   // 无成因 / no cause
    eCfgIllegal := 1,   // 组态非法：年月日、盘数或周期越域（故障级，与 bError 配对）/ illegal config, calendar, tray count or interval out of domain
    eTrayBad    := 2,   // 保养完成脉冲的托盘号越域已回钳（信息级）/ the tray number on the maintenance pulse was clamped, informational
    eNoDue      := 3    // 本月无到期盘（信息级）/ no tray is due this month, informational
);
END_TYPE

FUNCTION_BLOCK FB_DL_TrayMonthRotate
VAR_INPUT
    bEnable      : BOOL := TRUE;             // 使能，失能时掩码冻结保持末值 [-] / enable, the mask freezes and holds its last value when disabled
    bReset       : BOOL := FALSE;           // 复位上升沿清故障锁存与掩码 [-] / reset rising edge clears the fault latch and the mask
    nYear        : INT := 2026;              // 当前年份 [年]，域 2000..2100 / current year [year], domain 2000 to 2100
    nMonth       : INT := 1;                 // 当前月份 [月]，域 1..12 / current month [month], domain 1 to 12
    nDayOfMonth  : INT := 1;                 // 当月第几日 [日]，域 1..31 / day of month [day], domain 1 to 31
    nTrayCount   : INT := 12;                // 参与排程的托盘数 [个]，域 1..12 / scheduled tray count [count], domain 1 to 12
    nIntervalMonths : INT := 3;              // 保养周期 [月]，域 1..60 / maintenance interval [month], domain 1 to 60
    bMaintDone   : BOOL := FALSE;            // 保养完成脉冲，上升沿回写上次保养月 [-] / maintenance done pulse, the rising edge writes back the last maintenance month
    nMaintTray   : INT := 1;                 // 保养完成脉冲对应的托盘号 [盘号] / tray number carried by the maintenance pulse
END_VAR
VAR_IN_OUT
    anLastMaintMonth : ARRAY[1..12] OF INT;  // 逐托盘上次保养月（0 = 从未保养）[月]，引用型入参由调用方持有 / per tray last maintenance month, zero means never, reference parameter owned by the caller
END_VAR
VAR_OUTPUT
    wDueMask     : WORD := 16#0000;          // 到期托盘掩码，位 i-1 对应托盘 i [-] / due tray mask, bit i minus one maps to tray i
    nDueCount    : INT := 0;                 // 到期托盘数 [个] / due tray count
    nOverdueCount: INT := 0;                 // 超期托盘数（月差超周期）[个] / overdue tray count
    nPriTray     : INT := 0;                 // 本月轮换优先托盘号 [盘号] / rotation priority tray of the month
    bPriDue      : BOOL := FALSE;            // 优先托盘本月是否到期 [-] / whether the priority tray is due this month
    bDueToday    : BOOL := FALSE;            // 本月是否存在到期盘 [-] / whether any tray is due this month
    eCause       : E_DL_TmrCause := E_DL_TmrCause.eNone; // 成因出口 [枚举] / cause outlet [enum]
    bError       : BOOL := FALSE;            // 故障锁存标志 [-] / fault latch flag
END_VAR
VAR
    rtReset      : R_TRIG;                   // 复位沿检测，段 0 无条件刷新 / reset edge detector, refreshed unconditionally in segment zero
    rtMaint      : R_TRIG;                   // 保养完成沿检测，段 0 无条件刷新 / maintenance done edge detector, refreshed unconditionally in segment zero
    _eCause      : E_DL_TmrCause := E_DL_TmrCause.eNone;  // 内部成因 / internal cause
    _eFaultCause : E_DL_TmrCause := E_DL_TmrCause.eNone;  // 故障级成因，锁存至复位沿 / fault cause, latched until the reset edge
    _bFault      : BOOL := FALSE;            // 故障锁存位 [-] / fault latch bit
    _bInit       : BOOL := FALSE;            // 首扫初始化完成标志（R310）/ first scan initialisation flag
    _bCfgBad     : BOOL := FALSE;            // 组态非法判定 [-] / illegal configuration verdict
    _bTrayClamped: BOOL := FALSE;            // 回写托盘号被回钳 [-] / the write-back tray number was clamped
    _bDueBit     : BOOL := FALSE;            // 本条托盘到期判定 [-] / per tray due verdict
    _nUseCount   : INT := 0;                 // 钳定后的托盘数 [个] / clamped tray count
    _nInterval   : INT := 1;                 // 钳定后的保养周期 [月] / clamped maintenance interval [month]
    _nTray       : INT := 1;                 // 回写用托盘号（回钳 1..12）[盘号] / write-back tray number clamped one through twelve
    _nIdx        : INT := 1;                 // 托盘游标（1 起，回钳 1..12）[盘号] / tray cursor, one-based, clamped one through twelve
    _nLast       : INT := 0;                 // 本条托盘上次保养月 [月] / last maintenance month of the tray [month]
    _nElapsed    : INT := 0;                 // 距上次保养的月差 [月] / months since the last maintenance [month]
    _nPri        : INT := 1;                 // 轮换优先盘号工作值（1..12）[盘号] / rotation priority working value, one through twelve [tray]
    _wMask       : WORD := 16#0000;          // 掩码工作字，先移位后置位（R327）/ mask working word, shift before setting
    _wBit        : WORD := 16#0001;          // 本条托盘位掩码 [-] / per tray bit mask
END_VAR
VAR CONSTANT
    DL_TMR_MAX       : INT := 12;            // 托盘容量与游标回钳上界 [个] / tray capacity and cursor clamp upper bound
    DL_TMR_INT_MIN   : INT := 1;             // 保养周期下限 [月] / maintenance interval floor [month]
    DL_TMR_INT_MAX   : INT := 60;            // 保养周期上限 [月] / maintenance interval ceiling [month]
    DL_TMR_YEAR_MIN  : INT := 2000;          // 年份下限 [年] / year floor [year]
    DL_TMR_YEAR_MAX  : INT := 2100;          // 年份上限 [年] / year ceiling [year]
    DL_TMR_DAY_MAX   : INT := 31;            // 月内最大天数 [日] / maximum days within a month [day]
    DL_TMR_MONTHS    : INT := 12;            // 一周年月数，跨年回绕补齐用 [月] / months in a year for the wrap fill [month]
    DL_TMR_MASK_NONE : WORD := 16#0000;      // 空掩码常量 [-] / empty mask constant
    DL_TMR_MASK_ONE  : WORD := 16#0001;      // 单位位常量 [-] / single bit constant
END_VAR

// 段 0｜沿检测无条件周期刷新（禁入分支）/ segment 0, unconditional refresh of the edge detectors, never inside a branch
rtReset(CLK := bReset); // 复位沿无条件刷新 / unconditional refresh of the reset edge
rtMaint(CLK := bMaintDone); // 保养完成沿无条件刷新 / unconditional refresh of the maintenance edge

// 段 1｜首扫初始化（R310）/ segment 1, first scan initialisation
IF NOT _bInit THEN // 首扫一拍 / the very first scan
    _bInit := TRUE; // 置首扫完成标志 / raise the first scan flag
    _bFault := FALSE; // 故障锁存清零 / clear the fault latch
    _eCause := E_DL_TmrCause.eNone; // 信息级成因清零 / clear the informational cause
    _eFaultCause := E_DL_TmrCause.eNone; // 故障级成因清零 / clear the fault cause
    _wMask := DL_TMR_MASK_NONE; // 掩码清零 / clear the mask
END_IF

// 段 2｜复位沿作用域：清故障锁存 / 清掩码与统计（不改上次保养月表，属调用方资产）/ segment 2, reset edge scope
IF rtReset.Q THEN // 复位沿 / reset edge
    _bFault := FALSE; // 作用域一：清故障锁存 / scope one, clear the fault latch
    _eFaultCause := E_DL_TmrCause.eNone; // 作用域一：清故障级成因 / scope one, clear the fault cause
    _wMask := DL_TMR_MASK_NONE; // 作用域二：清到期掩码 / scope two, clear the due mask
    nDueCount := 0; // 作用域二：清到期计数 / scope two, clear the due count
    nOverdueCount := 0; // 作用域二：清超期计数 / scope two, clear the overdue count
END_IF

// 段 3｜组态域闸（R151 全覆盖）/ segment 3, configuration domain gate over every pin
_bCfgBad := FALSE; // 组态非法预置假 / preset the illegal configuration verdict to false
IF (nYear < DL_TMR_YEAR_MIN) OR (nYear > DL_TMR_YEAR_MAX) THEN // 年份越域 / year out of domain
    _bCfgBad := TRUE; // 判非法 / mark illegal
END_IF
IF (nMonth < 1) OR (nMonth > DL_TMR_MONTHS) THEN // 月份越域 / month out of domain
    _bCfgBad := TRUE; // 判非法 / mark illegal
END_IF
IF (nDayOfMonth < 1) OR (nDayOfMonth > DL_TMR_DAY_MAX) THEN // 当日序号越域 / day index out of domain
    _bCfgBad := TRUE; // 判非法 / mark illegal
END_IF
IF (nTrayCount < 1) OR (nTrayCount > DL_TMR_MAX) THEN // 托盘数越域 / tray count out of domain
    _bCfgBad := TRUE; // 判非法 / mark illegal
END_IF
IF (nIntervalMonths < DL_TMR_INT_MIN) OR (nIntervalMonths > DL_TMR_INT_MAX) THEN // 保养周期越域 / maintenance interval out of domain
    _bCfgBad := TRUE; // 判非法 / mark illegal
END_IF
IF _bCfgBad AND (NOT _bFault) THEN // 组态非法且未锁存 / illegal configuration and not yet latched
    _bFault := TRUE; // 置故障锁存 / raise the fault latch
    _eFaultCause := E_DL_TmrCause.eCfgIllegal; // 故障级成因 (R45 配对 bError) / fault grade cause paired with bError
END_IF
_nUseCount := nTrayCount; // 托盘数直通 / tray count passes through
IF _nUseCount < 1 THEN // 下越界 / below the lower bound
    _nUseCount := 1; // 回钳到 1 / clamp to one
ELSIF _nUseCount > DL_TMR_MAX THEN // 上越界 / above the upper bound
    _nUseCount := DL_TMR_MAX; // 回钳到容量上限 / clamp to the capacity ceiling
END_IF
_nInterval := nIntervalMonths; // 周期直通 / interval passes through
IF _nInterval < DL_TMR_INT_MIN THEN // 周期过小 / interval below the floor
    _nInterval := DL_TMR_INT_MIN; // 抬到下限 / raised to the floor
ELSIF _nInterval > DL_TMR_INT_MAX THEN // 周期过大 / interval above the ceiling
    _nInterval := DL_TMR_INT_MAX; // 压到上限 / pressed to the ceiling
END_IF

// 段 4｜保养完成回写：上升沿 + 托盘号回钳后写入上次保养月表 / segment 4, maintenance write-back on the rising edge with the tray number clamped
_bTrayClamped := FALSE; // 回钳标志预置假 / preset the clamp flag to false
IF rtMaint.Q THEN // 保养完成沿 / maintenance done edge
    _nTray := nMaintTray; // 托盘号直通 / tray number passes through
    IF _nTray < 1 THEN // 下越界 / below the lower bound
        _nTray := 1; // 回钳到 1 / clamp to one
        _bTrayClamped := TRUE; // 置回钳标志 / raise the clamp flag
    ELSIF _nTray > DL_TMR_MAX THEN // 上越界 / above the upper bound
        _nTray := DL_TMR_MAX; // 回钳到 12 / clamp to twelve
        _bTrayClamped := TRUE; // 置回钳标志 / raise the clamp flag
    END_IF
    anLastMaintMonth[_nTray] := nMonth; // 回写上次保养月，下标已回钳 1..12 / write back the last maintenance month with the index already clamped
END_IF

// 段 5｜逐盘到期判定与掩码打包 / segment 5, per tray due verdict and mask packing
_wMask := DL_TMR_MASK_NONE; // 掩码每拍清零重建 / the mask is rebuilt every scan
nDueCount := 0; // 到期计数清零 / clear the due count
nOverdueCount := 0; // 超期计数清零 / clear the overdue count
_nIdx := 1; // 游标自 1 起，上界由 _nUseCount 约束 / the cursor starts at one, bounded by the usable count
WHILE _nIdx <= _nUseCount DO // 循环上界为钳定后的托盘数，天然不越 12 / the loop bound is the clamped count, never beyond twelve
    _wBit := SHL(DL_TMR_MASK_ONE, _nIdx - 1); // 本条托盘位掩码，位移量 0..11 由数组边界与循环上界共同证明 / per tray bit mask, the shift zero through eleven is proven by the array and loop bounds
    _nLast := anLastMaintMonth[_nIdx]; // 上次保养月 / last maintenance month
    _bDueBit := FALSE; // 到期判定预置假 / preset the due verdict to false
    IF _nLast < 1 THEN // 从未保养 / never maintained
        _bDueBit := TRUE; // 立即到期 / due immediately
        nOverdueCount := nOverdueCount + 1; // 计入超期统计 / counted as overdue
    ELSE
        _nElapsed := nMonth - _nLast; // 月差 / month difference
        IF _nElapsed < 0 THEN // 跨年回绕 / year wrap
            _nElapsed := _nElapsed + DL_TMR_MONTHS; // 按月数补齐，仅覆盖一周年内 / filled by the months in a year, valid within one year
        END_IF
        IF _nElapsed >= _nInterval THEN // 达到周期 / the interval is reached
            _bDueBit := TRUE; // 判到期 / due verdict
            IF _nElapsed > _nInterval THEN // 超过周期 / beyond the interval
                nOverdueCount := nOverdueCount + 1; // 计入超期统计 / counted as overdue
            END_IF
        END_IF
    END_IF
    IF _bDueBit THEN // 本条托盘到期 / the tray is due
        _wMask := _wMask OR _wBit; // 置到期位 / set the due bit
        nDueCount := nDueCount + 1; // 到期计数递增 / increment the due count
    END_IF
    _nIdx := _nIdx + 1; // 游标递增 / increment the cursor
END_WHILE

// 段 6｜轮换优先盘号：按月份在托盘序列上轮转，除子为钳定后的托盘数 / segment 6, rotation priority tray with the clamped tray count as the divisor
_nPri := ((nMonth - 1) MOD _nUseCount) + 1; // 轮换公式，除子已证不小于 1 / rotation formula, divisor proven not below one
nPriTray := _nPri; // 优先盘号出口 / priority tray outlet
bPriDue := ((_wMask AND SHL(DL_TMR_MASK_ONE, _nPri - 1)) <> DL_TMR_MASK_NONE); // 优先盘是否到期，位移量 0..11 已证 / whether the priority tray is due, the shift zero through eleven is proven
bDueToday := nDueCount > 0; // 本月是否存在到期盘（挂状态量）/ whether any tray is due, a state quantity

// 段 7｜成因分派（固定优先级：故障 > 回钳 > 无到期 > 无成因）/ segment 7, cause dispatch with a fixed priority
IF _bFault THEN // 故障锁存优先 / the fault latch takes priority
    eCause := _eFaultCause; // 故障级成因锁存回放 / the fault cause is replayed from the latch
ELSIF _bTrayClamped THEN // 回写托盘号被回钳 / the write-back tray number was clamped
    eCause := E_DL_TmrCause.eTrayBad; // 信息级成因 / informational cause
ELSIF nDueCount < 1 THEN // 无到期盘 / no tray is due
    eCause := E_DL_TmrCause.eNoDue; // 信息级成因 / informational cause
ELSE
    eCause := E_DL_TmrCause.eNone; // 无成因 / no cause
END_IF

// 段 8｜统一出口 / segment 8, unified outlet
wDueMask := _wMask; // 到期掩码出口 / due mask outlet
bError := _bFault; // 故障标志与锁存位同源 / the fault flag shares the latch source
END_FUNCTION_BLOCK

(* ---- FB_DL_TunnelPasteurizerSeq.st ---- *)
(*==============================================================================
 * 组件名称 (Component)  : FB_DL_TunnelPasteurizerSeq
 * 所属子库 (Sublibrary) : DL_Process
 * 当前版本 (Version)    : 1.0.0
 * 兼容性   (Platform)   : CODESYS 3.5+ / TwinCAT 3 / 汇川 InoProShop / 施耐德 Machine Expert
 *                         仅依赖 Standard.library（TON / R_TRIG / ABS），零厂商私有库
 * 功能描述 (Function)   : 隧道式巴氏杀菌六态段序（保质期合规双联锁）：
 *                           ePreheat 预热：腔温升入杀菌带下沿（fTempPauSetC - fBandC）
 *                             → ePau；
 *                           ePau 杀菌：要求 ABS(fTempPau - fTempPauSetC) <= fBandC 且
 *                             tPauMin 驻留到时才放行 eCool；带外跌出**不退出 ePau 而冻结
 *                             驻留计时**（保守侧，TON IN 表达式派生）+ 记 eCause=eBandOut
 *                             （信息级每拍重算，回带即清）；
 *                           eCool 冷却：出口温降联锁 fTempCoo <= fCoolMaxC 才放行 eDone
 *                             （防烫瓶）；
 *                           进瓶无料（bBottleIn 长假）挂起不故障（不推进不算错）。
 * 接口     (Interface)  : 输入 bStart/bStop/bReset、fTempPau 杀菌区实测（℃）、fTempCoo
 *                         冷却区实测（℃）、fTempPauSetC 杀菌设定（℃）、fBandC 温度带
 *                         半宽（℃）、fCoolMaxC 出口允许最高温（℃）、tPauMin 杀菌段最短
 *                         驻留、tPreheatMin 预热最短时长、fVconvMmS 网链速度（mm/s）、
 *                         bBottleIn/bBottleOut 进出口光电；输出 ePhase 六态、bPauInBand
 *                         带内指示、相指示 BOOL 组、bDone、eCause、bError。
 * 边界     (Boundary)   : ① **属主边界（写死）：本件只做三温区段序推进与双联锁判定，不
 *                         驱动加热阀/风机/网链变频**（网链速度仅作诊断输入不内环控制）。
 *                         ② 六态 CASE + ELSE 兜底 eFault（R6）；TON 段 0 无条件刷新，
 *                         IN 由当前相与带内判据派生（带外冻结驻留，R188 自派生式）。
 *                         ③ 非有限温度 → eFault eCause=eNoData（分码，R190 归因唯一）。
 *                         ④ 组态闸：fBandC<=0、fCoolMaxC<=0、tPauMin<=T#0S、
 *                         tPreheatMin<=T#0S → 锁存 eFault eCfgIllegal。
 *                         ⑤ eCause 语义分层：eBandOut 为信息级（带内每拍重算清除）、
 *                         eNoData/eCfgIllegal 为故障级锁存（解除沿 = bReset 上升沿）。
 *                         ⑥ 温度带判定浮点全用 <= / >= 比较，禁 = 判等（R28）。
 *                         ⑦ 零全局耦合（无 GVL / VAR_EXTERNAL / 物理地址）。
 * 分工声明 (Scope)      : 与 `FB_DL_KilnSoakHoldCtrl` 类烧成件分域：巴杀温带驻留 ≠ 烧成
 *                         保温；与干燥段序件分域：出口温降联锁为食品保质期语义。
 * 来源标签 (Source Tag) : T2-2 ◐（LBP 工艺分层只借杀菌/冷却段序分类事实，双联锁实现自研）
 * 码表     (Codes)      : 本件不占用任何全局数字码位。出口为 ENUM 六态 + BOOL 组 +
 *                         ENUM 成因；数字码位待主控收口阶段统一派号。
 * 红线自检 (Redline)    : R1 ✓ 零 GVL/VAR_EXTERNAL ｜ R2 ✓ 零 %I/%Q/%M ｜ R3 ✓ 纯 IEC 61131-3
 *                         R4 ✓ 带冻结 TON 派生 + 非有限分码 + 组态闸 ｜ R5 ✓ 声明逐行同行双语注释
 *                         R6 ✓ 六态 CASE 含 ELSE ｜ R7 ✓ 两 TON/两 R_TRIG 段 0 无条件刷新
 * 修订历史 (Revision)   : 2026-11-20  v1.0.0  R48 首版（批次 4 · 序号 19）
 *                         验收向量：预热入带 → ePau；带外跌出驻留冻结不退出；tPauMin 到
 *                         + 带内 → eCool；出口超温禁 done；无料挂起不故障。
 *==============================================================================*)

TYPE E_DL_TpsPhase :
(
    eIdle    := 0,    // 待机 / Idle
    ePreheat := 10,   // 预热相 / Preheat phase
    ePau     := 20,   // 杀菌驻留相 / Pasteurization dwell phase
    eCool    := 30,   // 冷却相 / Cooling phase
    eDone    := 40,   // 程序完成 / Sequence done
    eFault   := 90    // 故障（等复位）/ Fault, awaiting reset
);
END_TYPE

TYPE E_DL_TpsCause :
(
    eNone       := 0,   // 无异常 / No anomaly
    eCfgIllegal := 1,   // 组态非法 / Illegal configuration
    eNoData     := 2,   // 温度非有限（故障级锁存）/ Non-finite temperature, latched
    eBandOut    := 3    // 杀菌带外（信息级，带内自动清除）/ Band dropout, informational
);
END_TYPE

FUNCTION_BLOCK FB_DL_TunnelPasteurizerSeq
VAR_INPUT
    bStart      : BOOL := FALSE;    // 启动沿（eIdle 入预热相） [-] / Start edge
    bStop       : BOOL := FALSE;    // 中止（任一相回 eIdle，不记故障） [-] / Abort to idle
    bReset      : BOOL := FALSE;    // 复位，上升沿清全部锁存（R311） [-] / Reset, rising edge clears all latches
    fTempPau    : LREAL := 0.0;     // 杀菌区实测温度 [℃] / Pasteurization zone temperature [degC]
    fTempCoo    : LREAL := 0.0;     // 冷却区实测温度 [℃] / Cooling zone temperature [degC]
    fTempPauSetC: LREAL := 72.0;    // 杀菌设定温度，域 > 0 [℃] / Pasteurization setpoint [degC]
    fBandC      : LREAL := 1.0;     // 杀菌温度带半宽，域 > 0 [℃] / Band half-width [degC]
    fCoolMaxC   : LREAL := 40.0;    // 出口允许最高温（温降联锁），域 > 0 [℃] / Outlet max temperature [degC]
    tPauMin     : TIME := T#10M;    // 杀菌段最短驻留，域 > T#0S [ms] / Minimum pasteurization dwell [ms]
    tPreheatMin : TIME := T#5M;     // 预热段最短时长，域 > T#0S [ms] / Minimum preheat duration [ms]
    fVconvMmS   : LREAL := 0.0;     // 网链速度（诊断输入，不内环控制） [mm/s] / Conveyor speed, diagnostic only [mm/s]
    bBottleIn   : BOOL := FALSE;    // 进瓶光电（长假期挂起不故障） [-] / Infeed photo-eye
    bBottleOut  : BOOL := FALSE;    // 出瓶光电（冷却段放行参考） [-] / Discharge photo-eye
END_VAR
VAR_OUTPUT
    ePhase     : E_DL_TpsPhase;     // 当前相出口 [-] / Present phase outlet
    bPauInBand : BOOL;              // 杀菌温度带内指示 [-] / In-band indicator
    bPreheatActive: BOOL;           // 预热相指示 [-] / Preheat indicator
    bPauActive : BOOL;              // 杀菌相指示 [-] / Pasteurization indicator
    bCoolActive: BOOL;              // 冷却相指示 [-] / Cooling indicator
    bDone      : BOOL;              // 程序完成（eDone 驻留指示） [-] / Done indicator
    eCause     : E_DL_TpsCause;     // 成因出口（信息级/故障级分层，头注释⑤） / Cause outlet
    bError     : BOOL;              // 故障标志 [-] / Error flag
END_VAR
VAR
    _eState  : E_DL_TpsPhase := E_DL_TpsPhase.eIdle;   // 内部相（CASE 唯一写入目标） / Internal phase
    _eCause  : E_DL_TpsCause := E_DL_TpsCause.eNone;   // 成因锁存量 / Latched cause
    _bFault  : BOOL;             // 故障锁存位（解除沿 = bReset 上升沿） / Latched fault bit
    _bInBand : BOOL;             // 当拍杀菌带内判据 [-] / In-band this scan
    _bNonFin : BOOL;             // 温度非有限当拍量 [-] / Non-finite temperature this scan
    _bCfgBad : BOOL;             // 组态非法当拍量 [-] / Illegal configuration this scan
    _bBusyPrev: BOOL;            // 上拍运行快照（bDone 迁出用） / Busy snapshot
    tonPreheat: TON;             // 预热最短时长定时器，段 0 无条件调用 / Preheat minimum timer
    tonPauMin : TON;             // 杀菌驻留计时定时器（带内派生 IN），段 0 无条件调用 / Pasteurization dwell timer
    rtStart   : R_TRIG;          // 启动沿实例，段 0 无条件调用 / Start edge instance
    rtReset   : R_TRIG;          // 复位沿实例，段 0 无条件调用 / Reset edge instance
END_VAR
VAR CONSTANT
    DL_TPS_ZERO : LREAL := 0.0;    // 非有限差值判零基准 [-] / Non-finite difference zero base
END_VAR

(* —— 段 0：非有限判 + 组态闸 + 两 TON 两沿无条件周期刷新 —— *)
_bNonFin := (fTempPau <> fTempPau) OR ((fTempPau - fTempPau) <> DL_TPS_ZERO)
         OR (fTempCoo <> fTempCoo) OR ((fTempCoo - fTempCoo) <> DL_TPS_ZERO);   // 双区温度非有限（R245） / Non-finite zone temperatures
_bCfgBad := (fBandC <= 0.0) OR (fCoolMaxC <= 0.0) OR (fTempPauSetC <= 0.0)
         OR (tPauMin <= T#0S) OR (tPreheatMin <= T#0S);     // 组态域闸 / Configuration gate
rtStart(CLK := bStart);                                     // 启动沿，每拍必调 / Start edge, every scan
rtReset(CLK := bReset);                                     // 复位沿，每拍必调 / Reset edge, every scan

(* —— 段 1：带内判据 + 驻留 TON 派生刷新（带外冻结驻留计时） —— *)
_bInBand := (NOT _bNonFin) AND (ABS(fTempPau - fTempPauSetC) <= fBandC);   // 杀菌带内（容差比较，禁 =） / In-band test
tonPreheat(IN := (_eState = E_DL_TpsPhase.ePreheat), PT := tPreheatMin);   // 预热最短计时（进相计时，出相自复位） / Preheat timer
tonPauMin(IN := (_eState = E_DL_TpsPhase.ePau) AND _bInBand, PT := tPauMin);   // 杀菌驻留计时（带外冻结，保守侧） / Dwell timer, band-gated

(* —— 段 2：单拍量预清零（锁存量 _eState/_eCause/_bFault 不入清单，R107） —— *)
bPreheatActive := FALSE;                                    // 预热相指示预清 / Preheat preset
bPauActive := FALSE;                                        // 杀菌相指示预清 / Pau preset
bCoolActive := FALSE;                                       // 冷却相指示预清 / Cool preset
bDone := FALSE;                                             // 完成指示预清 / Done preset
bError := FALSE;                                            // 故障标志预清（R45 配对） / Error preset

(* —— 段 3：组态闸入故障 —— *)
IF _bCfgBad AND (NOT _bFault) THEN
    _bFault := TRUE;                                        // 锁存 / Latch
    _eCause := E_DL_TpsCause.eCfgIllegal;                   // 归因：组态非法 / Cause: illegal config
    _eState := E_DL_TpsPhase.eFault;                        // 入故障相 / Enter fault
END_IF

(* —— 段 4：迁出链（bStop 优先不记故障；bReset 清全部锁存 R311） —— *)
IF bStop AND (_eState <> E_DL_TpsPhase.eIdle) THEN
    IF _eState = E_DL_TpsPhase.eFault THEN
        _bFault := FALSE;                                   // 停机优先清故障 / Stop wins over fault
        _eCause := E_DL_TpsCause.eNone;                     // 清成因 / Clear cause
    END_IF
    _eState := E_DL_TpsPhase.eIdle;                         // 回待机 / Back to idle
END_IF
IF rtReset.Q THEN
    _bFault := FALSE;                                       // 清故障锁存（R311） / Clear fault latch
    _eCause := E_DL_TpsCause.eNone;                         // 清成因 / Clear cause
    _eState := E_DL_TpsPhase.eIdle;                         // 回待机 / Back to idle
END_IF

(* —— 段 5：六态段序（只在无故障时推进；非有限 → 故障分码 eNoData） —— *)
IF (NOT _bFault) AND (NOT _bCfgBad) AND (NOT bStop) THEN
    IF _bNonFin AND (_eState <> E_DL_TpsPhase.eIdle) AND (_eState <> E_DL_TpsPhase.eDone) THEN
        _bFault := TRUE;                                    // 运行相温度非有限：故障锁存（规格③） / Non-finite in running phase
        _eCause := E_DL_TpsCause.eNoData;                   // 归因分码：无有效数据 / Cause: no data
        _eState := E_DL_TpsPhase.eFault;                    // 入故障相 / Enter fault
    ELSE
        CASE _eState OF

        E_DL_TpsPhase.eIdle:
            IF rtStart.Q THEN
                _eState := E_DL_TpsPhase.ePreheat;          // 启动沿入预热相 / Start edge enters preheat
            END_IF

        E_DL_TpsPhase.ePreheat:
            IF tonPreheat.Q AND (fTempPau >= (fTempPauSetC - fBandC)) THEN
                _eState := E_DL_TpsPhase.ePau;              // 预热到时 ∧ 温升入带下沿：进杀菌相 / Preheat done and in lower band
            END_IF

        E_DL_TpsPhase.ePau:
            IF _bInBand THEN
                _eCause := E_DL_TpsCause.eNone;             // 回带：清除信息级带外码（信息级每拍重算） / Back in band: clear info code
            ELSE
                _eCause := E_DL_TpsCause.eBandOut;          // 带外跌出：记信息级码，不退出不故障（规格③） / Band out: info code only
            END_IF
            IF tonPauMin.Q AND _bInBand THEN
                _eState := E_DL_TpsPhase.eCool;             // 驻留到时 ∧ 带内：放行冷却相 / Dwell done and in band: proceed
            END_IF

        E_DL_TpsPhase.eCool:
            _eCause := E_DL_TpsCause.eNone;                 // 冷却相清除信息级码 / Clear info code in cooling
            IF (fTempCoo <= fCoolMaxC) AND bBottleOut THEN
                _eState := E_DL_TpsPhase.eDone;             // 出口温降联锁 ∧ 出瓶：进完成相（防烫瓶） / Outlet cool enough with bottle out
            END_IF

        E_DL_TpsPhase.eDone:
            ;                                               // 完成相驻留：由 bReset / bStop 迁出 / Held, exits via reset or stop

        E_DL_TpsPhase.eFault:
            ;                                               // 故障相驻留：由迁出链处理 / Held by exit chain

        ELSE
            _eCause := E_DL_TpsCause.eCfgIllegal;           // 非法相位兜底归因 / Illegal phase cause
            _bFault := TRUE;                                // 锁存 / Latch
            _eState := E_DL_TpsPhase.eFault;                // 强拉故障相 / Force fault

        END_CASE
    END_IF
END_IF

(* —— 段 6：完成脉冲（由"运行→eDone"沿派生，单拍，R34 两段式） —— *)
IF _bBusyPrev AND (_eState = E_DL_TpsPhase.eDone) THEN
    bDone := TRUE;                                          // 程序完成单拍指示 / Done pulse
END_IF
_bBusyPrev := (_eState <> E_DL_TpsPhase.eIdle)
          AND (_eState <> E_DL_TpsPhase.eDone)
          AND (_eState <> E_DL_TpsPhase.eFault);            // 运行中快照（本拍末） / Busy snapshot at body end

(* —— 段 7：出口单点映射（相指示与相别同源，R191） —— *)
bPreheatActive := (_eState = E_DL_TpsPhase.ePreheat);       // 预热相指示 / Preheat indicator
bPauActive := (_eState = E_DL_TpsPhase.ePau);               // 杀菌相指示 / Pau indicator
bCoolActive := (_eState = E_DL_TpsPhase.eCool);             // 冷却相指示 / Cool indicator
IF _eState = E_DL_TpsPhase.eDone THEN
    bDone := TRUE;                                          // 完成相驻留期保持指示（R191） / Done held while resident
END_IF
bPauInBand := (_eState = E_DL_TpsPhase.ePau) AND _bInBand;   // 带内指示（仅杀菌相有意义） / In-band indicator
ePhase := _eState;                                          // 当前相出口 / Present phase outlet
eCause := _eCause;                                          // 成因出口 / Cause outlet
bError := _bFault OR _bCfgBad;                              // 故障标志 = 锁存或组态非法 / Error flag

END_FUNCTION_BLOCK

(* ---- FB_DL_UtilitiesLoadMgr.st ---- *)
(*==============================================================================
 * 组件名称 (Component)  : FB_DL_UtilitiesLoadMgr
 * 所属子库 (Sublibrary) : DL_Process
 * 前缀     (Prefix)     : FB_DL_
 * 当前版本 (Version)    : 1.0.0
 * 兼容性   (Platform)   : CODESYS 3.5 / TwinCAT 3 / 汇川 InoProShop / Schneider
 *                         Machine Expert；纯 IEC 61131-3（第 3 版），
 *                         仅依赖标准库 TON / R_TRIG / ABS / MAX / MIN，零厂商方言
 * 作者     (Author)     : 道莅代码库 · PLC编程专家（R31）
 * 开源溯源 (Origin)     : 多机按需投切负荷分配公开工艺语义（行业池，空压机/
 *                         冷冻机通用），轮值均衡借鉴本库 DutyStandbyRotation
 *                         思想（累计运行时长排序，零代码复制），道莅
 *                         clean-room 防御性实现，未复制任何外部源码行
 * 功能描述 (Function)   : 多机按需投切负荷分配件（空压机/冷冻机通用，不出
 *                         冷机专用变体）。加权平均负载对照回差双阈值
 *                         （启动阈高于停止阈防振荡）定增/减台数；投切按
 *                         累计运行时长均衡轮值；台数变更经驻留时间抑制。
 *                         仅指令与反馈持续矛盾置故障级，其余全部信息级。
 * 码位     (Codes)      : 16#0005_00B7 信息级：组态非法不投切、负载非有限
 *                                      权重归零、台数/阈值钳位（不置 bError）
 *                         16#0005_00B8 故障级：指令与反馈持续矛盾（锁存，
 *                                      bRst 复位沿为可达解除路径）
 *                         16#0005_00B9~00BB 保留未启用（码表与实现对齐）
 * 边界防错 (Boundary)   : 1 uMachCnt 为零或阈值倒置记组态码不投切；
 *                         2 非有限负载该机权重归零后均值重算防除零；
 *                         3 越界输出逐位清零；
 *                         4 TON/R_TRIG 实例每拍无条件刷新；
 *                         5 手动模式（bAuto=FALSE）冻结投切保持现状。
 * 修订历史 (Revision)   : 2026-11-18 v1.0.0 首版入库（R31 · 阶段三 · 序 17）
 *==============================================================================*)

(*==============================================================================
 * 功能块: FB_DL_UtilitiesLoadMgr
 * 调用约定: 每个扫描周期无条件调用一次；负载与运行反馈经引脚数组注入。
 *==============================================================================*)
FUNCTION_BLOCK FB_DL_UtilitiesLoadMgr
VAR_INPUT
    afLoad  : ARRAY[1..8] OF REAL;    // 各机负载率 [百分数] / Per-machine load rate [%]
    abFb    : ARRAY[1..8] OF BOOL;    // 各机运行反馈（可增引脚，矛盾判据用）/ Per-machine running feedback, added pin
    uMachCnt: UINT := 8;              // 机组台数 [台]，合法域 1..8 / Machine count, valid 1..8
    fStartTh: REAL := 80.0;           // 投切启动阈 [百分数]，须高于停止阈 / Start threshold [%], above stop
    fStopTh : REAL := 50.0;           // 投切停止阈 [百分数] / Stop threshold [%]
    uMinRun : UINT := 1;              // 最少运行台数 [台] / Minimum running count
    uMaxRun : UINT := 8;              // 最多运行台数 [台] / Maximum running count
    bAuto   : BOOL := FALSE;          // 自动模式 / Auto mode
    tDwell  : TIME := T#60S;          // 台数变更驻留 [毫秒] / Switching dwell [ms]
    tFbConf : TIME := T#10S;          // 反馈矛盾确认时长 [毫秒]（可增引脚）/ Feedback mismatch confirm [ms], added pin
    bRst    : BOOL := FALSE;          // 故障复位沿（可增引脚）/ Fault reset edge, added pin
END_VAR
VAR_OUTPUT
    abRun   : ARRAY[1..8] OF BOOL;    // 各机运行指令 / Per-machine run command
    uRunCnt : UINT;                   // 当前运行台数 [台] / Current running count
    bError  : BOOL;                   // 故障标志，与故障级码配对（R45）/ Fault flag paired with fault codes
    uErrorId: UDINT;                  // 错误码，0 = 无错 / Error code, 0 = none
END_VAR
VAR
    rTrigRst: R_TRIG;                 // 复位沿检测，每拍无条件刷新 / Reset edge detector, refreshed every scan
    tonDwell: TON;                    // 驻留计时，每拍无条件刷新 / Dwell timer, refreshed every scan
    tonFb   : TON;                    // 反馈矛盾确认计时，每拍无条件刷新 / Feedback mismatch timer
    i       : INT;                    // 逐机循环索引 / Per-machine loop index
    j       : INT;                    // 轮值选择内层索引 / Rotation inner loop index
    uCntEff : INT;                    // 钳位后有效台数 [台]，INT 域 / Effective clamped count, INT domain
    uMinEff : INT;                    // 钳位后最少台数 [台] / Effective minimum count
    uMaxEff : INT;                    // 钳位后最多台数 [台] / Effective maximum count
    nRunNow : INT;                    // 本拍运行台数 [台] / Running count this scan
    nValid  : INT;                    // 有限负载数 [台] / Finite load count
    fSum    : REAL;                   // 有限负载和 [百分数] / Finite load sum [%]
    fAvg    : REAL;                   // 加权平均负载 [百分数] / Weighted average load [%]
    bCfgOk  : BOOL;                   // 组态合法标志 / Configuration legality flag
    bAddReq : BOOL;                   // 增台请求 / Add request
    bSubReq : BOOL;                   // 减台请求 / Sub request
    bPickOk : BOOL;                   // 轮值选机成功 / Rotation pick success
    nSel    : INT;                    // 轮值选中下标 / Rotation selected index
    uTicksLo: UDINT;                  // 轮值最短累计时标 [拍] / Rotation shortest tick count
    auTicks : ARRAY[1..8] OF UDINT;   // 各机累计运行时标 [拍] / Per-machine run tick counters
    bAnyMis : BOOL;                   // 任一机指令反馈矛盾 / Any command-feedback mismatch
    bClamp  : BOOL;                   // 本拍钳位信息 / Clamp info this scan
    bDwellGo: BOOL;                   // 驻留期满许可投切 / Dwell elapsed permit
    xDwellRst: BOOL;                  // 投切拍单拍断驻留输入 / One-scan dwell input break after switch
    bFirst  : BOOL := TRUE;           // 首扫标志 / First-scan flag
END_VAR
VAR CONSTANT
    DL_ULD_MACH_MAX: INT  := 8;       // 台数上限 [台] / Machine count upper bound
    DL_ULD_FIN     : REAL := 1.0E30;  // REAL 有限幅值判界 / REAL finiteness magnitude bound
END_VAR

// ---- 段 1｜边沿与定时器实例无条件周期刷新（红线：禁入条件分支）----------------
rTrigRst(CLK := bRst);                                // 复位沿检测 / Reset edge detection
tonDwell(IN := ((NOT bFirst) AND (NOT xDwellRst)), PT := tDwell); // 驻留计时，投切拍断输入 / Dwell timing, broken on switch scan
tonFb(IN := bAnyMis, PT := tFbConf);                  // 矛盾确认计时 / Mismatch confirm timing

// ---- 段 2｜台数与阈值钳位（统一 INT 域）----------------------------------------
uCntEff := MIN(UINT_TO_INT(uMachCnt), DL_ULD_MACH_MAX); // 台数钳上限 / Clamp count to upper bound
uCntEff := MAX(uCntEff, 1);                           // 下限保 1 / Floor at 1
uMaxEff := MIN(UINT_TO_INT(uMaxRun), uCntEff);        // 最多台数钳到台数内 / Clamp max into count
uMaxEff := MAX(uMaxEff, 0);                           // 非负 / Non-negative
uMinEff := MIN(UINT_TO_INT(uMinRun), uMaxEff);        // 最少台数不超最多 / Min not above max
uMinEff := MAX(uMinEff, 0);                           // 非负 / Non-negative
bCfgOk := (uCntEff >= 1) AND (fStartTh > fStopTh) AND (fStartTh = fStartTh)
      AND (fStopTh = fStopTh) AND (ABS(fStartTh) < DL_ULD_FIN) AND (ABS(fStopTh) < DL_ULD_FIN); // 组态合法性 / Configuration legality
bClamp := (UINT_TO_INT(uMachCnt) > DL_ULD_MACH_MAX) OR (fStartTh <= fStopTh); // 钳位/倒置信息 / Clamp or inversion info

// ---- 段 3｜首拍与越界清位（越界逐位清零）----------------------------------------
IF bFirst THEN
    FOR i := 1 TO DL_ULD_MACH_MAX DO
        abRun[i] := FALSE;                            // 首拍全 FALSE / First scan all FALSE
        auTicks[i] := 0;                              // 时标清零 / Ticks cleared
    END_FOR
    bFirst := FALSE;                                  // 清首扫标志 / Clear first-scan flag
END_IF

// ---- 段 4｜负载有效性掩码与加权平均（非有限权重归零后均值重算防除零）------------
nValid := 0;                                          // 有效数清零 / Clear valid count
fSum := 0.0;                                          // 和清零 / Clear sum
FOR i := 1 TO uCntEff DO
    IF (afLoad[i] = afLoad[i]) AND (ABS(afLoad[i]) < DL_ULD_FIN) THEN
        nValid := nValid + 1;                         // 有效负载计数 / Count finite load
        fSum := fSum + afLoad[i];                     // 累加有效负载 / Accumulate finite load
    END_IF
END_FOR
IF nValid > 0 THEN
    fAvg := fSum / UDINT_TO_REAL(INT_TO_UDINT(nValid)); // 均值，分母已验正 / Average, denominator verified
ELSE
    fAvg := 0.0;                                      // 全无效确定值 / Deterministic fallback
END_IF

// ---- 段 5｜运行台数统计与时标累计 ------------------------------------------------
nRunNow := 0;                                         // 台数清零 / Clear count
FOR i := 1 TO uCntEff DO
    IF abRun[i] THEN
        nRunNow := nRunNow + 1;                       // 统计运行台数 / Count running machines
        auTicks[i] := auTicks[i] + 1;                 // 运行时标累计（轮值均衡基准）/ Run ticks accumulate
    END_IF
END_FOR

// ---- 段 6｜投切决策（组态非法或非自动冻结投切；驻留期满许可）--------------------
bDwellGo := tonDwell.Q;                               // 驻留期满 / Dwell elapsed
bAddReq := bCfgOk AND bAuto AND bDwellGo AND (fAvg > fStartTh) AND (nRunNow < uMaxEff); // 增台请求 / Add request
bSubReq := bCfgOk AND bAuto AND bDwellGo AND (fAvg < fStopTh) AND (nRunNow > uMinEff); // 减台请求 / Sub request
IF bAddReq THEN
    bPickOk := FALSE;                                 // 选机标志先清 / Clear pick flag
    uTicksLo := 16#FFFFFFFF;                          // 最短时标预置满 / Preset shortest ticks full
    FOR j := 1 TO uCntEff DO
        IF (NOT abRun[j]) AND (auTicks[j] < uTicksLo) THEN
            uTicksLo := auTicks[j];                   // 更新最短时标 / Update shortest ticks
            nSel := j;                                // 记录选中下标 / Record selected index
            bPickOk := TRUE;                          // 选机成功 / Pick success
        END_IF
    END_FOR
    IF bPickOk THEN
        abRun[nSel] := TRUE;                          // 投入最短时标停运机 / Start shortest-tick idle machine
        xDwellRst := TRUE;                            // 投切拍断驻留输入重置计时 / Break dwell input on switch scan
    END_IF
ELSIF bSubReq THEN
    bPickOk := FALSE;                                 // 选机标志先清 / Clear pick flag
    uTicksLo := 0;                                    // 最长时标预置零 / Preset longest ticks zero
    FOR j := 1 TO uCntEff DO
        IF abRun[j] AND (auTicks[j] >= uTicksLo) THEN
            uTicksLo := auTicks[j];                   // 更新最长时标 / Update longest ticks
            nSel := j;                                // 记录选中下标 / Record selected index
            bPickOk := TRUE;                          // 选机成功 / Pick success
        END_IF
    END_FOR
    IF bPickOk THEN
        abRun[nSel] := FALSE;                         // 停运最长时标运行机 / Stop longest-tick running machine
        xDwellRst := TRUE;                            // 投切拍断驻留输入重置计时 / Break dwell input on switch scan
    END_IF
END_IF

// ---- 段 7｜指令反馈矛盾监视与故障锁存 --------------------------------------------
bAnyMis := FALSE;                                     // 矛盾标志先清 / Clear mismatch flag
FOR i := 1 TO uCntEff DO
    IF abRun[i] AND (NOT abFb[i]) THEN
        bAnyMis := TRUE;                              // 指令真反馈假矛盾 / Command true feedback false
    END_IF
END_FOR
IF rTrigRst.Q THEN
    bAnyMis := FALSE;                                 // 复位清矛盾路径 / Reset clears mismatch path
END_IF

// ---- 段 8｜输出台数与错误码装配 --------------------------------------------------
nRunNow := 0;                                         // 重统计输出台数 / Recount running
FOR i := 1 TO DL_ULD_MACH_MAX DO
    IF i > uCntEff THEN
        abRun[i] := FALSE;                            // 越界逐位清零 / Out-of-range bits cleared
    END_IF
    IF abRun[i] THEN
        nRunNow := nRunNow + 1;                       // 输出台数统计 / Count output running
    END_IF
END_FOR
uRunCnt := INT_TO_UINT(nRunNow);                      // 台数输出 / Count output
IF tonFb.Q THEN
    bError   := TRUE;                                 // 指令反馈持续矛盾锁故障 / Persistent mismatch latches fault
    uErrorId := 16#0005_00B8;                         // 码位：矛盾持续 / Code: persistent mismatch
ELSIF (NOT bCfgOk) OR bClamp OR (nValid = 0) THEN
    bError   := FALSE;                                // 信息级不置故障 / Info never sets fault
    uErrorId := 16#0005_00B7;                         // 信息级：组态/非有限/钳位 / Info: config or non-finite
ELSE
    bError   := FALSE;                                // 无错清标志 / Clear fault flag
    uErrorId := 16#0000_0000;                         // 无码 / No code
END_IF

// ---- 段 9｜单拍标志收尾 ----------------------------------------------------------
xDwellRst := FALSE;                                   // 断输入请求仅当拍有效 / Break request is single scan
END_FUNCTION_BLOCK

(* ---- FB_DL_VacCupRingCtrl.st ---- *)
(*
    FB_DL_VacCupRingCtrl —— 多吸盘组分档拾放
    ------------------------------------------------------------------
    分类      : DL_Process / Handling
    前缀      : FB_DL_
    版本      : 1.0.0
    溯源      : 多吸盘拾放为公开搬运工程结构（成组吸附 → 确认 → 分组释放）；
                逐通道确认、少吸失败判据、分组释放相、降级放行、错误分级与码位 100% 自有；
                单个真空发生器仍归设备层（本件不内联真空发生器控制）；
                clean-room 重写，未复制任何闭源厂商源码
    平台      : 纯 IEC 61131-3，CODESYS V3.5+ / TwinCAT 3 / InoProShop 通用
    作者      : 道莅代码库 · PLC编程专家（R19）
    ------------------------------------------------------------------
    功能说明  : 一组（1~8 个）真空吸盘的拾放控制：逐通道吸附确认、吸盘数不足时判拾取
                失败（安全侧：少吸的料上轴会在加速时掉落）、可选降级放行（少吸但达最低
                要求）、分组释放（先外圈后内圈，防料被甩）。
                核心防御：① 吸盘数越界、最少需吸附数大于总数、真空门限非负或超物理可达——
                   三类参数错即故障级 0308 并撤销全部阀输出，绝不索引数组；
                ② 逐通道判据 = 到位开关闭合 **且** 真空度低于门限，两者同时成立才算到位
                   （只看开关会漏掉管路微漏，只看数值会被单点噪声骗过）；
                ③ 真空值非有限按「未到位」处理并置故障级 0309，绝不当成到位；
                ④ 确认时间到而到位数不足即锁存拾取失败，保持吸附（掉料比保持更危险）；
                ⑤ 降级放行必须显式允许（bAllowDegrade）且达到最低吸盘数；
                ⑥ 分组释放两相，相内不改吸附判据；⑦ CASE 含 ELSE 兜底回 eIdle 并撤阀。
                职责边界：真空发生器/喷射器的单机控制归设备层件，本件只做组级工艺编排。
    错误码    : 16#0005_01D8 降级放行（少吸但达最低要求）/ 拾取计数饱和——信息级，正常防御
                16#0005_01D9 预留禁用（信息级，不得挪用）
                16#0005_0308 吸盘数或真空门限参数非法——故障级，阀输出全部撤销
                16#0005_0309 吸附确认失败（到位数不足 / 真空值非有限 / 确认超时）——故障级，锁存并保持吸附
                16#0005_030A 状态机落 ELSE 兜底（非法状态）——故障级，回 eIdle 并撤销阀输出（用途固定，不得改作他用）
    码位总账  : 16#0005_01D8 用 / 16#0005_01D9 预留 ｜ 16#0005_0308 用 / 16#0005_0309 用 / 16#0005_030A 用
    状态机    : E_DL_VacRingState（eIdle / ePicking / eHolding / eReleasing / eDegraded / eFault）六态，
                CASE 含 ELSE 兜底，ELSE 回 eIdle 并撤销全部阀输出。
    采样约定  : fbTrigReset / fbTrigPick / fbTrigRelease 与 fbConfirm / fbSettle 五个实例在本体首部
                无条件刷新，绝不放入 IF 或 CASE（按段断输入是本族高危点）；
                释放两相各自计时：fbConfirm 覆盖「外圈已释放」，fbSettle 覆盖「内圈已释放」。
    修订记录  : 2026-11-16 v1.0.0 首次入库（R19）
*)

(*
    枚举 : E_DL_VacRingState —— 吸盘组拾放状态（本文件为全库唯一属主）
*)
TYPE E_DL_VacRingState :
(
    eIdle      := 0,                          // 空闲：无吸附无动作 / idle, nothing held and no action
    ePicking   := 1,                          // 拾取中：等待吸附确认 / picking, waiting for the vacuum confirmation
    eHolding   := 2,                          // 保持中：全部吸盘确认到位 / holding, every cup confirmed
    eReleasing := 3,                          // 释放中：两相分组释放 / releasing, two phase grouped release
    eDegraded  := 4,                          // 降级保持：少吸但达最低要求 / degraded hold, fewer cups but above the minimum
    eFault     := 5                           // 故障：参数错或拾取失败 / fault, parameter error or pick failure
);
END_TYPE

FUNCTION_BLOCK FB_DL_VacCupRingCtrl
VAR_INPUT
    bEnable            : BOOL;                // 使能，FALSE 撤销所有阀输出 / enable, FALSE withdraws every valve output
    bReset             : BOOL;                // 复位，上升沿清故障与降级锁存 / reset, rising edge clears the faults and the degraded latch
    bCmdPick           : BOOL;                // 拾取命令（上升沿启动）/ pick command, rising edge starts it
    bCmdRelease        : BOOL;                // 释放命令（上升沿启动）/ release command, rising edge starts it
    auVacuumOk         : ARRAY[0..7] OF BOOL; // 各吸盘真空到位开关 / vacuum reached switch per cup
    afVacuum           : ARRAY[0..7] OF REAL; // 各吸盘真空度（负值）[kPa]，范围 -101.3~0.0 / vacuum level per cup, negative [kPa], range -101.3~0.0
    uCupCount          : UINT := 4;           // 有效吸盘数 [个]，范围 1~8 / valid cup count [cup], range 1~8
    uMinCupsRequired   : UINT := 4;           // 最少需吸附的吸盘数 [个]，范围 1~uCupCount / minimum cups to confirm [cup], range 1~uCupCount
    fVacMin            : REAL := -40.0;       // 真空度合格门限（负值，绝对值越大越紧）[kPa] / vacuum acceptance threshold, negative [kPa]
    tConfirmTime       : TIME := T#500MS;     // 吸附确认时间（亦作释放相时间）[ms]，范围 0~10000 / confirmation and release phase time [ms], range 0~10000
    bAllowDegrade      : BOOL := FALSE;       // TRUE = 允许少吸降级放行（须达最低要求）/ TRUE allows a degraded release above the minimum
    bReleaseOuterFirst : BOOL := TRUE;        // TRUE = 先释放偶数通道（视为外圈）/ TRUE releases the even channels first, treated as the outer ring
END_VAR
VAR_OUTPUT
    auValveOut         : ARRAY[0..7] OF BOOL; // 各吸盘真空阀输出（由上层映射到物理点）/ vacuum valve output per cup, mapped to physical points above
    bPicked            : BOOL;                // 已拾取（吸附确认通过）/ picked, the vacuum confirmation passed
    bReleased          : BOOL;                // 已释放完成 / released, the release finished
    uOkCups            : UINT;                // 当前确认到位的吸盘数 [个] / cups currently confirmed [cup]
    bDegraded          : BOOL;                // 降级运行中（少吸放行）/ running degraded with fewer cups
    bPickFailed        : BOOL;                // 拾取失败（锁存，需 bReset）/ pick failure, latched until reset
    uPickCount         : UDINT;               // 累计成功拾取次数，饱和 [次] / accumulated successful picks, saturating [times]
    eErr               : UDINT;               // 错误码，0=正常 / error id, 0=ok
    bError             : BOOL;               // 故障标志，eErr 为故障级时 TRUE / error flag, TRUE on fault-level eErr
END_VAR
VAR
    eState             : E_DL_VacRingState := eIdle; // 状态机当前态 / current state machine state
    fbTrigReset        : R_TRIG;              // 复位上升沿实例，本体首部无条件刷新 / reset edge instance, refreshed unconditionally
    fbTrigPick         : R_TRIG;              // 拾取命令沿实例，本体首部无条件刷新 / pick edge instance, refreshed unconditionally
    fbTrigRelease      : R_TRIG;              // 释放命令沿实例，本体首部无条件刷新 / release edge instance, refreshed unconditionally
    fbConfirm          : TON;                 // 吸附确认与释放第一相定时器，本体首部无条件刷新 / confirmation and first release phase timer, refreshed unconditionally
    fbSettle           : TON;                 // 释放第二相定时器，本体首部无条件刷新 / second release phase timer, refreshed unconditionally
    uIdx               : UINT;                // 通道扫描游标 [通道]，范围 0~7 / channel scan cursor [channel], range 0~7
    uOk                : UINT;                // 本拍到位的吸盘数 [个] / confirmed cups in this cycle [cup]
    uPhase             : UINT;                // 释放分组相号 [相]，0 = 外圈，1 = 内圈 / release phase index [phase], zero outer, one inner
    fVacMinEff         : REAL;                // 钳位后的真空门限 [kPa] / clamped vacuum threshold [kPa]
    bNonFinVac         : BOOL;                // 存在非有限真空值 / a non-finite vacuum value exists
    bGroupA            : BOOL;                // 本通道属于当前相要释放的分组 / this channel belongs to the group released in the current phase
    bInit              : BOOL := FALSE;       // 首扫标志，初值 FALSE，判据 NOT bInit / first-scan flag, initial FALSE, tested with NOT
    tConfirmEff        : TIME;                // 钳位后的确认时间（定时器 PT 前置收敛）[ms] / clamped confirmation time feeding the timers [ms]
END_VAR
VAR CONSTANT
    DL_VRC_CUP_MAX      : UINT := 8;          // 吸盘数上限 [个] / cup count upper bound [cup]
    DL_VRC_VAC_ABS_MAX  : REAL := 101.3;      // 真空物理上限（绝对值）[kPa] / absolute physical vacuum bound [kPa]
    DL_VRC_CNT_MAX      : UDINT := 16#FFFF_FFFE; // 拾取计数饱和值 [次] / pick counter saturation value [times]
    DL_VRC_DT_MAX       : TIME := T#10S;      // 确认时间上限 [ms] / confirmation time upper bound [ms]
    DL_FLOAT_EPS        : REAL := 1.0E-6;     // 浮点判等容差 [无量纲] / float equality tolerance [dimensionless]
    DL_VRC_INF_GUARD    : REAL := 1.0E38;     // 非有限幅值判定阈值 [无量纲] / non-finite magnitude guard [dimensionless]
    DL_VRC_TWO          : UINT := 2;          // 二值常量，内外圈分组用 [无量纲] / two constant used by the ring grouping
    DL_VRC_PHASE_ONE    : UINT := 1;          // 第二相相号 [相] / phase index of the second release
    DL_VRC_ZERO         : REAL := 0.0;        // 零值常量，避免裸字面量 [无量纲] / zero constant, avoids a bare literal [dimensionless]
    DL_VRC_CNT_ZERO     : UINT := 0;          // 无符号零常量 [无量纲] / unsigned zero constant [dimensionless]
END_VAR

// 段 1｜确认时间前置收敛（定时器 PT 的入参必须先合法）/ segment 1, clamp the confirmation time before the timers
tConfirmEff := tConfirmTime;                   // 取入参副本 / copy the input
IF tConfirmEff > DL_VRC_DT_MAX THEN
    tConfirmEff := DL_VRC_DT_MAX;              // 超上限钳到 10 s / clamp to ten seconds
END_IF
IF tConfirmEff < T#0S THEN
    tConfirmEff := T#0S;                       // 负时间无物理意义 / a negative time has no physical meaning
END_IF

// 段 2｜边沿与定时器实例无条件周期刷新（红线：严禁放入条件分支）/ segment 2, unconditional refresh
fbTrigReset(CLK := bReset);
fbTrigPick(CLK := bCmdPick);
fbTrigRelease(CLK := bCmdRelease);
fbConfirm(IN := (eState = ePicking) OR ((eState = eReleasing) AND (uPhase = DL_VRC_CNT_ZERO)), PT := tConfirmEff); // 拾取确认与释放第一相共用 / shared by the pick confirmation and the first release phase
fbSettle(IN := (eState = eReleasing) AND (uPhase >= DL_VRC_PHASE_ONE), PT := tConfirmEff);                          // 释放第二相计时 / times the second release phase

// 段 2｜输出与错误状态预置（bPicked / bPickFailed / uPickCount 为保持量）/ segment 2, preset outputs
eErr := 0;                                     // 预置无错误 / preset no error
bError := FALSE;                               // 预置无故障 / preset no fault
bReleased := FALSE;                            // 脉冲类标志先清 / clear the pulse style flags
uOkCups := DL_VRC_CNT_ZERO;                    // 到位数清零 / clear the confirmed cup count
uOk := DL_VRC_CNT_ZERO;                        // 到位数中间量清零 / clear the intermediate count
bNonFinVac := FALSE;                           // 预置无非有限真空值 / preset no non-finite vacuum
uPhase := DL_VRC_CNT_ZERO;                     // 相号复位 / reset the phase index
FOR uIdx := 0 TO DL_VRC_CUP_MAX - 1 DO
    auValveOut[uIdx] := FALSE;                 // 全部阀输出先撤销，再由状态逻辑按需置位 / clear every valve output, the state logic sets them again
END_FOR

// 段 3｜首扫初始化（唯一合法范式：初值 FALSE，判据 NOT bInit）/ segment 3, first-scan initialisation
IF NOT bInit THEN
    bPicked := FALSE;                          // 首扫未拾取 / not picked on the first scan
    bPickFailed := FALSE;                      // 首扫无拾取失败 / no pick failure on the first scan
    bDegraded := FALSE;                        // 首扫无降级 / not degraded on the first scan
    uPickCount := 0;                           // 拾取统计清零 / clear the pick statistics
    bInit := TRUE;                             // 首扫只做一次 / first scan runs once only
END_IF

// 段 4｜参数闸（三类参数错一律撤销阀输出，且绝不索引数组）/ segment 4, parameter gate
IF (uCupCount < 1) OR (uCupCount > DL_VRC_CUP_MAX) THEN
    eErr := 16#0005_0308;                      // 吸盘数越界故障码 / cup count out of range fault id
    bError := TRUE;                            // 置故障标志 / raise the error flag
    eState := eFault;                          // 落故障态 / enter the fault state
    RETURN;                                   // 故障级提前返回，阀输出已全撤 / early return, the valve outputs are already cleared
END_IF
IF (uMinCupsRequired < 1) OR (uMinCupsRequired > uCupCount) THEN
    eErr := 16#0005_0308;                      // 最少吸附数矛盾故障码 / contradictory minimum cup count fault id
    bError := TRUE;                            // 置故障标志 / raise the error flag
    eState := eFault;                          // 落故障态 / enter the fault state
    RETURN;                                   // 故障级提前返回 / early return on fault
END_IF
IF (fVacMin <> fVacMin) OR (fVacMin >= DL_VRC_ZERO) OR (ABS(fVacMin) > DL_VRC_VAC_ABS_MAX) THEN
    eErr := 16#0005_0308;                      // 真空门限非负或不可达故障码 / the vacuum threshold is non-negative or unreachable
    bError := TRUE;                            // 置故障标志 / raise the error flag
    eState := eFault;                          // 落故障态 / enter the fault state
    RETURN;                                   // 故障级提前返回 / early return on fault
END_IF

// 段 5｜真空门限域钳位（确认时间已在段 1 收敛）/ segment 5, threshold clamp, the confirmation time was clamped in segment 1
fVacMinEff := MAX(fVacMin, -DL_VRC_VAC_ABS_MAX); // 门限绝对值收敛到物理可达 [kPa] / converge the threshold into the physical range [kPa]

// 段 6｜使能闸：失能撤销所有阀输出 / segment 6, enable gate
IF NOT bEnable THEN
    eState := eIdle;                           // 回空闲态 / back to idle
    bPicked := FALSE;                          // 不计已拾取 / not picked
    bDegraded := FALSE;                        // 撤降级 / drop the degraded flag
    RETURN;                                   // 失能即出口，阀输出已全撤 / disabled is the exit, the outputs are already cleared
END_IF

// 段 7｜复位沿：清故障与降级锁存（不改变吸附状态）/ segment 7, reset clears the latches
IF fbTrigReset.Q THEN
    bPickFailed := FALSE;                      // 清拾取失败锁存 / clear the pick failure latch
    bDegraded := FALSE;                        // 清降级锁存 / clear the degraded latch
    bPicked := FALSE;                          // 清已拾取标志 / clear the picked flag
    IF eState = eFault THEN
        eState := eIdle;                       // 故障态由复位退出 / a reset leaves the fault state
    END_IF
END_IF

// 段 8｜逐通道吸附确认（到位开关与真空度必须同时成立）/ segment 8, per channel confirmation
FOR uIdx := 0 TO uCupCount - 1 DO
    IF (afVacuum[uIdx] <> afVacuum[uIdx]) OR (afVacuum[uIdx] > DL_VRC_INF_GUARD) OR (afVacuum[uIdx] < -DL_VRC_INF_GUARD) THEN
        bNonFinVac := TRUE;                    // 非有限真空值：按未到位处理，绝不当成到位 / a non-finite value counts as not confirmed, never as confirmed
    ELSIF auVacuumOk[uIdx] AND (afVacuum[uIdx] <= fVacMinEff) THEN
        uOk := uOk + 1;                        // 开关与数值同时成立才计入 / both the switch and the level must agree
    END_IF
END_FOR
uOkCups := uOk;                                // 发布到位吸盘数 [个] / publish the confirmed cup count [cup]

// 段 9｜状态机（含 ELSE 兜底）/ segment 9, state machine with ELSE fallback
CASE eState OF
    eIdle:
        bPicked := FALSE;                      // 空闲不计已拾取 / idle is not picked
        IF fbTrigPick.Q THEN
            eState := ePicking;                // 拾取沿进入拾取中 / a pick edge enters the picking state
        ELSIF fbTrigRelease.Q THEN
            uPhase := DL_VRC_CNT_ZERO;         // 释放从第一相开始 / the release starts in the first phase
            eState := eReleasing;              // 直接进入释放（空手释放用于清管）/ entering release with nothing held is allowed to purge
        END_IF

    ePicking:
        FOR uIdx := 0 TO uCupCount - 1 DO
            auValveOut[uIdx] := TRUE;          // 拾取相全部吸盘抽真空 / every cup is evacuated in the picking phase
        END_FOR
        IF bNonFinVac THEN
            eErr := 16#0005_0309;              // 真空值非有限故障码 / non-finite vacuum fault id
            bError := TRUE;                    // 置故障标志 / raise the error flag
            bPickFailed := TRUE;               // 锁存拾取失败 / latch the pick failure
            eState := eFault;                  // 落故障态（保持吸附，掉料更危险）/ the fault state keeps the vacuum, dropping the load is worse
        ELSIF uOk >= uCupCount THEN
            bPicked := TRUE;                   // 全部到位即拾取成功 / every cup confirmed means a successful pick
            IF uPickCount < DL_VRC_CNT_MAX THEN
                uPickCount := uPickCount + 1;  // 饱和累计拾取次数 / saturating pick counter
            END_IF
            eState := eHolding;                // 进入保持态 / enter the holding state
        ELSIF (uOk >= uMinCupsRequired) AND bAllowDegrade THEN
            bDegraded := TRUE;                  // 少吸但达最低要求且显式允许：降级放行 / fewer cups but above the minimum and explicitly allowed
            bPicked := TRUE;                    // 降级也算拾取（工艺已允许）/ a degraded pick still counts, the process allowed it
            eErr := 16#0005_01D8;               // 信息级：降级放行 / info level, released in a degraded mode
            eState := eDegraded;                // 进入降级保持态 / enter the degraded holding state
        ELSIF fbConfirm.Q THEN
            eErr := 16#0005_0309;               // 确认超时仍未到位故障码 / the confirmation timed out short of the minimum
            bError := TRUE;                     // 置故障标志 / raise the error flag
            bPickFailed := TRUE;                // 锁存拾取失败（安全侧：少吸的料上轴会掉落）/ latch the failure, carrying a partial load would drop it during acceleration
            eState := eFault;                   // 落故障态并保持吸附 / enter the fault state and keep the vacuum
        END_IF

    eHolding:
        FOR uIdx := 0 TO uCupCount - 1 DO
            auValveOut[uIdx] := TRUE;          // 保持相持续抽真空 / the holding phase keeps the vacuum
        END_FOR
        IF fbTrigRelease.Q THEN
            uPhase := DL_VRC_CNT_ZERO;         // 释放从第一相开始 / start with the first phase
            eState := eReleasing;              // 进入释放相 / enter the release phase
        END_IF

    eDegraded:
        FOR uIdx := 0 TO uCupCount - 1 DO
            auValveOut[uIdx] := TRUE;          // 降级保持同样保持真空 / the degraded hold keeps the vacuum as well
        END_FOR
        bDegraded := TRUE;                      // 持续发布降级标志 / keep publishing the degraded flag
        IF fbTrigRelease.Q THEN
            uPhase := DL_VRC_CNT_ZERO;         // 释放从第一相开始 / start with the first phase
            eState := eReleasing;              // 进入释放相 / enter the release phase
        END_IF

    eReleasing:
        // 段 10｜分组释放：第一相放外圈（偶数通道），第二相放内圈 / segment 10, two phase grouped release
        FOR uIdx := 0 TO uCupCount - 1 DO
            IF uPhase = DL_VRC_CNT_ZERO THEN
                IF bReleaseOuterFirst THEN
                    bGroupA := (uIdx MOD DL_VRC_TWO) = DL_VRC_CNT_ZERO; // 偶数通道为外圈 / the even channels form the outer ring
                ELSE
                    bGroupA := (uIdx MOD DL_VRC_TWO) <> DL_VRC_CNT_ZERO; // 奇数通道为外圈 / the odd channels form the outer ring
                END_IF
                auValveOut[uIdx] := NOT bGroupA; // 第一相只放外圈，其余继续抽真空 / only the outer ring is released in the first phase
            ELSE
                auValveOut[uIdx] := FALSE;      // 第二相全部释放 / everything is released in the second phase
            END_IF
        END_FOR
        IF (uPhase = DL_VRC_CNT_ZERO) AND fbConfirm.Q THEN
            uPhase := DL_VRC_PHASE_ONE;         // 第一相到时进入第二相 / the first phase elapses into the second
        ELSIF (uPhase >= DL_VRC_PHASE_ONE) AND fbSettle.Q THEN
            bReleased := TRUE;                  // 释放完成单周期脉冲 / the release completed, a single-cycle pulse
            bPicked := FALSE;                   // 清已拾取 / clear the picked flag
            bDegraded := FALSE;                 // 清降级 / clear the degraded flag
            uPhase := DL_VRC_CNT_ZERO;          // 相号复位 / reset the phase index
            eState := eIdle;                    // 回空闲态 / back to idle
        END_IF

    eFault:
        // 段 11｜故障态：参数错时阀已全撤；拾取失败时保持吸附 / segment 11, the fault state keeps the vacuum after a pick failure
        IF bPickFailed THEN
            FOR uIdx := 0 TO uCupCount - 1 DO
                auValveOut[uIdx] := auVacuumOk[uIdx]; // 保持已确认的通道，未确认的不再抽（避免持续漏气补压）/ keep the confirmed cups, stop evacuating those that never confirm
            END_FOR
        END_IF

ELSE
    eErr := 16#0005_030A;                       // 故障级：非法状态兜底（用途固定）/ fault level, illegal state fallback, the purpose is fixed
    bError := TRUE;                             // 置故障标志 / raise the error flag
    eState := eIdle;                            // 回空闲态 / fall back to idle
    FOR uIdx := 0 TO DL_VRC_CUP_MAX - 1 DO
        auValveOut[uIdx] := FALSE;              // 兜底时撤销全部阀输出 / withdraw every valve output on the fallback path
    END_FOR
END_CASE
END_FUNCTION_BLOCK
